(* IEC 61131-3 sources: PortalRobot/Portal_robot/Device/application/FB (part 2) *)

(* ---- FB_AXIS_GROUP.st ---- *)
FUNCTION_BLOCK FB_AXIS_GROUP
VAR_INPUT
	FaultRequest : ST_AXIS_GROUP_FAULT_REQUEST; // Единый контракт диагностической инъекции
	xResetPermit : BOOL; // Общий сброс разрешён ручным режимом и остановленной ячейкой
	xAxesPowered : BOOL; // Питанием физических осей владеют FB_AXIS; группа только наблюдает готовность
	lrVelocityOverride : LREAL; // Live override скорости групповых движений, 0.001..1.0
END_VAR
VAR_OUTPUT
	FaultStatus : ST_FAULT_INJECTION_STATUS; // Состояние инжектора для HMI
END_VAR
VAR
	// Внутренние исполняемые булевые переменные
	xEnable      : BOOL; // Импульс включения группы
	xDisable     : BOOL; // Импульс отключения группы
	xReset       : BOOL; // Импульс сброса ошибок
	xResetMC     : BOOL; // Выполняется сброс SoftMotion
	xMoveDirect  : BOOL; // Выполняется прямое перемещение
	xMoveLinear  : BOOL; // Выполняется линейное перемещение
	xStopCmd     : BOOL; // Выполняется остановка
	xHaltCmd     : BOOL; // Выполняется плавная остановка
	lrAppliedVelocityOverride : LREAL; // Коэффициент после защитного ограничения PLC
	xVelocityOverrideEnable : BOOL; // Запись live override разрешена только в рабочих состояниях без MC_GroupStop
	xFaultAllowed : BOOL; // Безопасные условия тестового запуска

	iPrevStep : E_AXIS_GROUP_STATE; // Предыдущий шаг автомата

	// Для таймера шага
	tonStepTimeout   : TON; // Таймер превышения времени шага
	xStepTimeout     : BOOL; // Время шага превышено
	xStepChanged     : BOOL; // Шаг изменился в текущем цикле
	xStepTimerEnable : BOOL; // Разрешение таймера шага
	xStepInitialized : BOOL; // Предыдущий шаг инициализирован

	// Для удержания предупреждений
    tpWarningHold : TP; // Удержание предупреждения для отображения
    xWarningPulse : BOOL; // Импульс нового предупреждения

	// ФБ группы осей
	fbReadStatus   : MC_GroupReadStatus; // Чтение состояния группы
	fbReadError    : MC_GroupReadError; // Чтение активной ошибки группы
	fbReadPosition : MC_GroupReadActualPosition; // Чтение текущей позиции группы
	fbGroupEnable  : MC_GroupEnable; // Включение группы
	fbGroupDisable : MC_GroupDisable; // Отключение группы
	fbGroupReset   : MC_GroupReset; // Сброс ошибок группы
	fbGroupSetOverride : MC_GroupSetOverride; // Live override активного и следующего движения группы

	fbMoveDirect : MC_MoveDirectAbsolute; // Прямое абсолютное перемещение
	fbMoveLinear : MC_MoveLinearAbsolute; // Линейное абсолютное перемещение
	fbFaultInjector : FB_AXIS_GROUP_FAULT_INJECTOR; // Изолированная инъекция библиотечной ошибки

	fbGroupHalt : MC_GroupHalt; // Плавная остановка группы
	fbGroupStop : MC_GroupStop; // Остановка группы

	stPosition : SMC_POS_REF; // Текущая позиция группы

	// Триггеры на команды
    rtEnable        : R_TRIG; // Фронт команды включения
    rtDisable       : R_TRIG; // Фронт команды отключения
	rtEnablePower   : R_TRIG; // Фронт запроса питания
    rtResetAllError : R_TRIG; // Фронт команды сброса
    rtMoveDirect    : R_TRIG; // Фронт прямого перемещения
    rtMoveLinear    : R_TRIG; // Фронт линейного перемещения
	rtStopCmd       : R_TRIG; // Фронт команды остановки
	rtHaltCmd       : R_TRIG; // Фронт плавной остановки

END_VAR
VAR_IN_OUT
	AxisGroup : AXIS_GROUP_REF_SM3; // Ссылка на группу осей SoftMotion
	GroupData : ST_AXIS_GROUP; // Команды, статусы и диагностика группы
END_VAR

VAR CONSTANT
	// ==================================================
    // Логические ошибки группы
    // ==================================================
	LOG_STEP_TIMEOUT             : DWORD := 1; // Превышено время шага
	LOG_INVALID_STATE            : DWORD := 2; // Неизвестный шаг автомата
	LOG_POWER_PERMIT_READY       : DWORD := 4; // Нет разрешения питания в готовности
	LOG_POWER_PERMIT_LOST_DIRECT : DWORD := 8; // Разрешение питания снято при движении
	// ==================================================
    // Ошибки блоков движения группы
    // ==================================================
	MOTION_ERR_ENABLE        : DWORD := 1; // Ошибка включения группы
	MOTION_ERR_DISABLE       : DWORD := 4; // Ошибка отключения группы
	MOTION_ERR_RESET         : DWORD := 8; // Ошибка сброса группы
	MOTION_ERR_MOVE_DIRECT   : DWORD := 16; // Ошибка прямого перемещения
	MOTION_ERR_MOVE_LINEAR   : DWORD := 32; // Ошибка линейного перемещения
	MOTION_ERR_HALT          : DWORD := 64; // Ошибка плавной остановки
	MOTION_ERR_STOP          : DWORD := 128; // Ошибка остановки
	MOTION_ERR_READ_POSITION : DWORD := 256; // Ошибка чтения позиции
	MOTION_ERR_READ_STATUS   : DWORD := 512; // Ошибка чтения статуса
	MOTION_ERR_READ_GROUP_ERROR : DWORD := 1024; // Ошибка чтения кода ошибки группы
	MOTION_ERR_GROUP_ERROR_STOP : DWORD := 2048; // Группа SoftMotion находится в ErrorStop
	MOTION_ERR_SIMULATED        : DWORD := 4096; // Тестовая ошибка MC_MoveDirectAbsolute
	MOTION_ERR_OVERRIDE         : DWORD := 8192; // Ошибка MC_GroupSetOverride; бит 1 сохранён за legacy POWER_ERROR

	WRN_NO_POWER_PERMIT       : UINT := 1; // Нет разрешения питания
	WRN_MOVE_COMMAND_CONFLICT : UINT := 2; // Одновременно заданы два типа движения
	WRN_GLOBAL_ERROR_ACTIVE   : UINT := 3; // Сброс отклонён из-за глобальной ошибки
	WRN_MOTION_ERROR_ACTIVE   : UINT := 4; // Сброс отклонён из-за активной Motion-ошибки
	WRN_RESET_VERIFY_TIMEOUT  : UINT := 5; // Не получено подтверждение сброса за допустимое время
	WRN_GROUP_ERROR_AFTER_RESET : UINT := 6; // Группа осталась в ErrorStop после сброса
	WRN_GROUP_RESET_ERROR     : UINT := 7; // MC_GroupReset завершился ошибкой
	WRN_GROUP_RESET_TIMEOUT   : UINT := 8; // Превышено время выполнения MC_GroupReset
	WRN_SIM_ERROR_NOT_ALLOWED : UINT := 9; // Тестовая ошибка запрещена текущим состоянием группы
END_VAR

// --- BEGIN IMPLEMENTATION ---

// Коэффициент симуляции не изменяет динамику группы осей робота.
lrAppliedVelocityOverride := MAX(0.001, MIN(1.0, lrVelocityOverride));

// =============================================================================
// 1. Добить предупреждения и ошибки
// 2. Сделать логирование ошибок и шагов
// 3. Сделать необходимые сигналы статусов
// =============================================================================

// =============================================================================
// 1. Одноцикловые сигналы
// =============================================================================
xWarningPulse := FALSE;

GroupData.Diag.xStepChanged := FALSE;
GroupData.Error.dwLogicalErrorNew := DWORD#0;
GroupData.Error.dwMotionErrorNew := DWORD#0;

// =============================================================================
// 2. Фронты команд
// =============================================================================
rtDisable(CLK := GroupData.Command.xDisable);
rtEnablePower(CLK := GroupData.Command.xPowerEnable);
rtResetAllError(CLK := GroupData.Command.xReset);
rtMoveDirect(CLK := GroupData.Command.xMoveDirect);
rtMoveLinear(CLK := GroupData.Command.xMoveLinear);
rtHaltCmd(CLK := GroupData.Command.xHaltCmd);
rtStopCmd(CLK := GroupData.Command.xStopCmd);

// =============================================================================
// 3. Чтение состояния группы и координат
// =============================================================================
fbReadStatus(
    Enable    := TRUE,
    AxisGroup := AxisGroup
);

fbReadError(
    Enable    := TRUE,
    AxisGroup := AxisGroup
);

fbReadPosition(
    AxisGroup   := AxisGroup,
    Enable      := TRUE,
    CoordSystem := SMC_COORD_SYSTEM.MCS
);

IF fbReadPosition.Valid THEN
	stPosition := fbReadPosition.Position;
    GroupData.Status.ActualX := fbReadPosition.Position.c.X;
    GroupData.Status.ActualY := fbReadPosition.Position.c.Y;
    GroupData.Status.ActualZ := fbReadPosition.Position.c.Z;
END_IF;
GroupData.Status.xPositionValid := fbReadPosition.Valid AND NOT fbReadPosition.Error;

// =============================================================================
// 4. Текущий статус ошибок
// =============================================================================
GroupData.Status.xGroupError :=
    fbReadStatus.Error
    OR fbReadStatus.GroupErrorStop
    OR (GroupData.Error.dwMotionErrorLatched <> DWORD#0);

GroupData.Status.xLogicalError :=
    GroupData.Error.dwLogicalErrorLatched <> DWORD#0;

GroupData.Status.xLocalError :=
    GroupData.Status.xGroupError
    OR GroupData.Status.xLogicalError;

// Тестовый Motion-FB запускается только в неподвижной готовой группе.
xFaultAllowed := fbReadStatus.Valid
	AND fbReadStatus.GroupStandby
	AND (GroupData.Diag.iStep = E_AXIS_GROUP_STATE.READY)
	AND NOT GroupData.Status.xLocalError
	AND NOT GroupData.Command.xGlobalError
	AND NOT GroupData.Command.xMoveDirect
	AND NOT GroupData.Command.xMoveLinear;

fbFaultInjector(
	Request := FaultRequest,
	xOwnerAllowed := xFaultAllowed,
	xReset := GroupData.Command.xReset,
	Position := stPosition,
	AxisGroup := AxisGroup
);
FaultStatus := fbFaultInjector.Status;

IF fbFaultInjector.Status.xRejected THEN
	GroupData.Diag.sWarningText := 'Simulated SM3 error is not allowed';
	GroupData.Diag.stWarning.uiCode := WRN_SIM_ERROR_NOT_ALLOWED;
	GroupData.Diag.stWarning.udiSequence := GroupData.Diag.stWarning.udiSequence + UDINT#1;
	IF GroupData.Diag.stWarning.udiSequence = UDINT#0 THEN
		GroupData.Diag.stWarning.udiSequence := UDINT#1;
	END_IF;
	xWarningPulse := TRUE;
END_IF;

// =============================================================================
// 5. Команды Motion FB по умолчанию
// =============================================================================
xEnable := FALSE;
xDisable := FALSE;
xResetMC := FALSE;
xMoveDirect := FALSE;
xMoveLinear := FALSE;
xStopCmd := FALSE;
xHaltCmd := FALSE;

// =============================================================================
// 6. Машина состояний
// =============================================================================
CASE GroupData.Diag.iStep OF

    // -------------------------------------------------------------------------
    E_AXIS_GROUP_STATE.DISABLED:
    // -------------------------------------------------------------------------
        GroupData.Diag.sStepName := 'DISABLED';
        GroupData.Diag.tStepPreset := T#0S;
        GroupData.Diag.iPowerMode := E_AXIS_GROUP_POWER_MODE.OFF;

        IF GroupData.Command.xGlobalError
           OR GroupData.Status.xLocalError THEN

            GroupData.Diag.iStep := E_AXIS_GROUP_STATE.ERROR;

        ELSIF rtEnablePower.Q AND NOT GroupData.Command.xPowerPermit THEN
            GroupData.Diag.sWarningText := 'Power permit is not active';
            GroupData.Diag.stWarning.uiCode := WRN_NO_POWER_PERMIT;
            GroupData.Diag.stWarning.udiSequence := GroupData.Diag.stWarning.udiSequence + UDINT#1;
            IF GroupData.Diag.stWarning.udiSequence = UDINT#0 THEN
                GroupData.Diag.stWarning.udiSequence := UDINT#1;
            END_IF;
            xWarningPulse := TRUE;

		ELSIF fbReadStatus.Valid AND fbReadStatus.GroupStandby THEN
			// MC_GroupReset всегда возвращает группу в GroupStandby. Если питание
			// запрошено, используем это состояние без повторного MC_GroupEnable;
			// иначе сначала синхронизируем группу с программным шагом DISABLED.
			IF rtEnablePower.Q THEN
				GroupData.Diag.iStep := E_AXIS_GROUP_STATE.ENABLING_POWER;
			ELSE
				GroupData.Diag.iStep := E_AXIS_GROUP_STATE.DISABLING_GROUP;
			END_IF;

        ELSIF rtEnablePower.Q THEN
            GroupData.Diag.iStep := E_AXIS_GROUP_STATE.ENABLING_POWER;
        END_IF;

    // -------------------------------------------------------------------------
    E_AXIS_GROUP_STATE.ENABLING_POWER:
    // -------------------------------------------------------------------------
        GroupData.Diag.sStepName := 'ENABLING_POWER';
        GroupData.Diag.tStepPreset := GroupData.Timeouts.tPowerTimeout;
        GroupData.Diag.iPowerMode := E_AXIS_GROUP_POWER_MODE.ON;

        IF fbReadStatus.GroupErrorStop THEN

            GroupData.Diag.iStep := E_AXIS_GROUP_STATE.ERROR;

        ELSIF NOT GroupData.Command.xPowerPermit
           OR GroupData.Command.xGlobalError THEN

            GroupData.Diag.iStep := E_AXIS_GROUP_STATE.DISABLING_POWER;

        ELSIF xStepTimeout THEN
            GroupData.Error.dwLogicalErrorNew :=
                GroupData.Error.dwLogicalErrorNew
                OR LOG_STEP_TIMEOUT;

            GroupData.Diag.iStep := E_AXIS_GROUP_STATE.DISABLING_POWER;

		ELSIF xAxesPowered AND fbReadStatus.Valid THEN
			IF fbReadStatus.GroupStandby THEN
				GroupData.Diag.iStep := E_AXIS_GROUP_STATE.READY;
			ELSIF fbReadStatus.GroupDisabled THEN
				GroupData.Diag.iStep := E_AXIS_GROUP_STATE.ENABLING_GROUP;
			END_IF;
		END_IF;

    // -------------------------------------------------------------------------
    E_AXIS_GROUP_STATE.ENABLING_GROUP:
    // -------------------------------------------------------------------------
        GroupData.Diag.sStepName := 'ENABLING_GROUP';
        GroupData.Diag.tStepPreset := GroupData.Timeouts.tGroupTimeout;
        GroupData.Diag.iPowerMode := E_AXIS_GROUP_POWER_MODE.ON;

		// MC_GroupEnable допустим только из GroupDisabled. Execute формируется
		// исключительно на этом шаге: после перехода в GroupStandby он снимается,
		// чтобы новый фронт не вызвал MC_GroupEnable повторно после MC_GroupReset.
		xEnable := fbReadStatus.Valid AND fbReadStatus.GroupDisabled;

		IF fbReadStatus.GroupErrorStop THEN

            GroupData.Diag.iStep := E_AXIS_GROUP_STATE.ERROR;

		ELSIF fbReadStatus.Valid AND fbReadStatus.GroupStandby THEN

			GroupData.Diag.iStep := E_AXIS_GROUP_STATE.READY;

		ELSIF xEnable AND fbGroupEnable.Error THEN

			GroupData.Diag.iStep := E_AXIS_GROUP_STATE.ERROR;

        ELSIF NOT GroupData.Command.xPowerPermit
           OR GroupData.Command.xGlobalError THEN

            GroupData.Diag.iStep := E_AXIS_GROUP_STATE.DISABLING_GROUP;

        ELSIF xStepTimeout THEN
            GroupData.Error.dwLogicalErrorNew :=
                GroupData.Error.dwLogicalErrorNew
                OR LOG_STEP_TIMEOUT;

            GroupData.Diag.iStep := E_AXIS_GROUP_STATE.DISABLING_GROUP;

		END_IF;

    // -------------------------------------------------------------------------
    E_AXIS_GROUP_STATE.READY:
    // -------------------------------------------------------------------------
        GroupData.Diag.sStepName := 'READY';
        GroupData.Diag.tStepPreset := T#0S;
        GroupData.Diag.iPowerMode := E_AXIS_GROUP_POWER_MODE.ON;

		IF fbReadStatus.GroupErrorStop THEN
            GroupData.Diag.iStep := E_AXIS_GROUP_STATE.ERROR;

        ELSIF NOT GroupData.Command.xPowerPermit
           OR GroupData.Command.xGlobalError
           OR GroupData.Status.xLocalError
           OR rtDisable.Q THEN

            GroupData.Diag.iStep := E_AXIS_GROUP_STATE.DISABLING_GROUP;

        ELSIF rtMoveDirect.Q AND rtMoveLinear.Q THEN
            GroupData.Diag.sWarningText :=
                'MoveDirect and MoveLinear requested together';

            GroupData.Diag.stWarning.uiCode := WRN_MOVE_COMMAND_CONFLICT;
            GroupData.Diag.stWarning.udiSequence := GroupData.Diag.stWarning.udiSequence + UDINT#1;
            IF GroupData.Diag.stWarning.udiSequence = UDINT#0 THEN
                GroupData.Diag.stWarning.udiSequence := UDINT#1;
            END_IF;

            xWarningPulse := TRUE;

        ELSIF rtMoveDirect.Q THEN
            GroupData.Diag.iStep := E_AXIS_GROUP_STATE.MOVING_DIRECT;

        ELSIF rtMoveLinear.Q THEN
            GroupData.Diag.iStep := E_AXIS_GROUP_STATE.MOVING_LINEAR;
        END_IF;

    // -------------------------------------------------------------------------
    E_AXIS_GROUP_STATE.MOVING_DIRECT:
    // -------------------------------------------------------------------------
        GroupData.Diag.sStepName := 'MOVING_DIRECT';
        GroupData.Diag.tStepPreset := GroupData.Timeouts.tMoveTimeout;
        GroupData.Diag.iPowerMode := E_AXIS_GROUP_POWER_MODE.ON;

		xMoveDirect := TRUE;

        IF fbReadStatus.GroupErrorStop THEN
            GroupData.Diag.iStep := E_AXIS_GROUP_STATE.ERROR;

        ELSIF fbMoveDirect.Error THEN
            IF fbReadStatus.GroupMoving THEN
                GroupData.Diag.iStep := E_AXIS_GROUP_STATE.EMG_STOP;
            ELSE
                GroupData.Diag.iStep := E_AXIS_GROUP_STATE.ERROR;
            END_IF;

        ELSIF xStepTimeout THEN
            GroupData.Error.dwLogicalErrorNew :=
                GroupData.Error.dwLogicalErrorNew
                OR LOG_STEP_TIMEOUT;

            GroupData.Diag.iStep := E_AXIS_GROUP_STATE.EMG_STOP;

        ELSIF NOT GroupData.Command.xPowerPermit
           OR GroupData.Command.xGlobalError
           OR GroupData.Status.xLocalError
           OR rtStopCmd.Q THEN

            GroupData.Diag.iStep := E_AXIS_GROUP_STATE.EMG_STOP;

        ELSIF rtHaltCmd.Q THEN
            GroupData.Diag.iStep := E_AXIS_GROUP_STATE.HALT_STOP;

        ELSIF fbMoveDirect.Done
           AND fbReadStatus.GroupStandby THEN

            GroupData.Diag.iStep := E_AXIS_GROUP_STATE.READY;
        END_IF;

    // -------------------------------------------------------------------------
    E_AXIS_GROUP_STATE.HALT_STOP:
    // -------------------------------------------------------------------------
        GroupData.Diag.sStepName := 'HALT_STOP';
        GroupData.Diag.tStepPreset := GroupData.Timeouts.tHaltTimeout;
        GroupData.Diag.iPowerMode := E_AXIS_GROUP_POWER_MODE.ON;

		xHaltCmd := TRUE;

        IF fbReadStatus.GroupErrorStop THEN
            GroupData.Diag.iStep := E_AXIS_GROUP_STATE.ERROR;

        ELSIF fbGroupHalt.Error
           OR xStepTimeout
           OR NOT GroupData.Command.xPowerPermit
           OR GroupData.Command.xGlobalError
           OR GroupData.Status.xLocalError
           OR rtStopCmd.Q THEN

            IF xStepTimeout THEN
                GroupData.Error.dwLogicalErrorNew :=
                    GroupData.Error.dwLogicalErrorNew
                    OR LOG_STEP_TIMEOUT;
            END_IF;

            GroupData.Diag.iStep := E_AXIS_GROUP_STATE.EMG_STOP;

        ELSIF fbGroupHalt.Done
           AND fbReadStatus.GroupStandby THEN

            GroupData.Diag.iStep := E_AXIS_GROUP_STATE.READY;
        END_IF;

    // -------------------------------------------------------------------------
    E_AXIS_GROUP_STATE.EMG_STOP:
    // -------------------------------------------------------------------------
        GroupData.Diag.sStepName := 'STOPPING';
        GroupData.Diag.tStepPreset := GroupData.Timeouts.tStopTimeout;
        GroupData.Diag.iPowerMode := E_AXIS_GROUP_POWER_MODE.ON;

		xStopCmd := TRUE;

        IF fbReadStatus.GroupErrorStop
           OR fbGroupStop.Error THEN

            GroupData.Diag.iStep := E_AXIS_GROUP_STATE.ERROR;

        ELSIF xStepTimeout THEN
            GroupData.Error.dwLogicalErrorNew :=
                GroupData.Error.dwLogicalErrorNew
                OR LOG_STEP_TIMEOUT;

            GroupData.Diag.iStep := E_AXIS_GROUP_STATE.ERROR;

        ELSIF fbGroupStop.Done THEN
            GroupData.Diag.iStep := E_AXIS_GROUP_STATE.WAIT_STOP;
        END_IF;

    // -------------------------------------------------------------------------
    E_AXIS_GROUP_STATE.WAIT_STOP:
    // -------------------------------------------------------------------------
        GroupData.Diag.sStepName := 'WAIT_STOP';
        GroupData.Diag.tStepPreset := GroupData.Timeouts.tStopTimeout;
        GroupData.Diag.iPowerMode := E_AXIS_GROUP_POWER_MODE.ON;

		IF fbReadStatus.GroupErrorStop THEN
            GroupData.Diag.iStep := E_AXIS_GROUP_STATE.ERROR;

        ELSIF xStepTimeout THEN
            GroupData.Error.dwLogicalErrorNew :=
                GroupData.Error.dwLogicalErrorNew
                OR LOG_STEP_TIMEOUT;

            GroupData.Diag.iStep := E_AXIS_GROUP_STATE.ERROR;

		ELSIF fbReadStatus.GroupStandby THEN
			// Операторский Stop завершает только движение и сохраняет GroupStandby.
			// Отключение группы выполняется лишь по отдельному запросу питания/ошибке.
			IF GroupData.Command.xPowerPermit
			AND NOT GroupData.Command.xDisable
			AND NOT GroupData.Command.xGlobalError
			AND NOT GroupData.Status.xLocalError THEN
				GroupData.Diag.iStep := E_AXIS_GROUP_STATE.READY;
			ELSE
				GroupData.Diag.iStep := E_AXIS_GROUP_STATE.DISABLING_GROUP;
			END_IF;
		END_IF;

    // -------------------------------------------------------------------------
    E_AXIS_GROUP_STATE.DISABLING_GROUP:
    // -------------------------------------------------------------------------
        GroupData.Diag.sStepName := 'DISABLING_GROUP';
        GroupData.Diag.tStepPreset := GroupData.Timeouts.tGroupTimeout;
        GroupData.Diag.iPowerMode := E_AXIS_GROUP_POWER_MODE.ON;

		// MC_GroupDisable допустим только из GroupStandby.
		xDisable := fbReadStatus.Valid AND fbReadStatus.GroupStandby;

		IF fbReadStatus.GroupErrorStop THEN

            GroupData.Diag.iStep := E_AXIS_GROUP_STATE.ERROR;

		ELSIF fbReadStatus.Valid AND fbReadStatus.GroupDisabled THEN

			GroupData.Diag.iStep := E_AXIS_GROUP_STATE.DISABLING_POWER;

		ELSIF xDisable AND fbGroupDisable.Error THEN

			GroupData.Diag.iStep := E_AXIS_GROUP_STATE.ERROR;

        ELSIF xStepTimeout THEN
            GroupData.Error.dwLogicalErrorNew :=
                GroupData.Error.dwLogicalErrorNew
                OR LOG_STEP_TIMEOUT;

            GroupData.Diag.iStep := E_AXIS_GROUP_STATE.ERROR;

		ELSIF xDisable AND fbGroupDisable.Done
           AND fbReadStatus.GroupDisabled THEN

            GroupData.Diag.iStep := E_AXIS_GROUP_STATE.DISABLING_POWER;
        END_IF;

    // -------------------------------------------------------------------------
    E_AXIS_GROUP_STATE.DISABLING_POWER:
    // -------------------------------------------------------------------------
        GroupData.Diag.sStepName := 'DISABLING_POWER';
        GroupData.Diag.tStepPreset := GroupData.Timeouts.tPowerTimeout;
        GroupData.Diag.iPowerMode :=
            E_AXIS_GROUP_POWER_MODE.OFF_REQUEST;

        IF xStepTimeout THEN
            GroupData.Error.dwLogicalErrorNew :=
                GroupData.Error.dwLogicalErrorNew
                OR LOG_STEP_TIMEOUT;

            GroupData.Diag.iStep := E_AXIS_GROUP_STATE.ERROR;

        ELSIF NOT xAxesPowered THEN

            IF GroupData.Command.xGlobalError
               OR GroupData.Status.xLocalError
			   OR NOT GroupData.Command.xPowerPermit THEN

                GroupData.Diag.iStep := E_AXIS_GROUP_STATE.ERROR;
            ELSE
                GroupData.Diag.iStep := E_AXIS_GROUP_STATE.DISABLED;
            END_IF;
        END_IF;

    // -------------------------------------------------------------------------
    E_AXIS_GROUP_STATE.ERROR:
    // -------------------------------------------------------------------------
        GroupData.Diag.sStepName := 'ERROR';
        GroupData.Diag.tStepPreset := T#0S;

        GroupData.Diag.iPowerMode := E_AXIS_GROUP_POWER_MODE.OFF_REQUEST;

		IF rtResetAllError.Q AND xResetPermit THEN

            IF GroupData.Command.xGlobalError THEN
                GroupData.Diag.sWarningText :=
                    'Global error is still active';

                GroupData.Diag.stWarning.uiCode := WRN_GLOBAL_ERROR_ACTIVE;
                GroupData.Diag.stWarning.udiSequence := GroupData.Diag.stWarning.udiSequence + UDINT#1;
                IF GroupData.Diag.stWarning.udiSequence = UDINT#0 THEN
                    GroupData.Diag.stWarning.udiSequence := UDINT#1;
                END_IF;

                xWarningPulse := TRUE;

            ELSIF fbReadStatus.GroupErrorStop THEN
                    GroupData.Diag.iStep :=
                        E_AXIS_GROUP_STATE.RESETTING;

            ELSIF GroupData.Error.dwMotionErrorActive
                  <> DWORD#0 THEN

                GroupData.Diag.sWarningText :=
                    'Motion FB error is still active';

                GroupData.Diag.stWarning.uiCode := WRN_MOTION_ERROR_ACTIVE;
                GroupData.Diag.stWarning.udiSequence := GroupData.Diag.stWarning.udiSequence + UDINT#1;
                IF GroupData.Diag.stWarning.udiSequence = UDINT#0 THEN
                    GroupData.Diag.stWarning.udiSequence := UDINT#1;
                END_IF;

                xWarningPulse := TRUE;

            ELSE
                // Ошибка устранена — очищаем защёлки.
                GroupData.Error.dwLogicalErrorLatched := DWORD#0;
                GroupData.Error.dwMotionErrorLatched := DWORD#0;
                GroupData.Error.dwMotionErrorPrevious := DWORD#0;

				IF fbReadStatus.GroupStandby AND NOT xAxesPowered THEN
					GroupData.Diag.iStep :=
						E_AXIS_GROUP_STATE.DISABLING_GROUP;

				ELSIF fbReadStatus.GroupDisabled AND NOT xAxesPowered THEN
					GroupData.Diag.iStep :=
						E_AXIS_GROUP_STATE.DISABLED;

				ELSIF fbReadStatus.GroupDisabled THEN
					GroupData.Diag.iStep :=
						E_AXIS_GROUP_STATE.ENABLING_GROUP;

                ELSIF fbReadStatus.GroupStandby THEN
                    GroupData.Diag.iStep :=
                        E_AXIS_GROUP_STATE.READY;

                ELSE
                    GroupData.Diag.iStep :=
                        E_AXIS_GROUP_STATE.DISABLING_POWER;
                END_IF;
            END_IF;
        END_IF;

    // -------------------------------------------------------------------------
    E_AXIS_GROUP_STATE.RESETTING:
    // -------------------------------------------------------------------------
        GroupData.Diag.sStepName := 'RESETTING';
        GroupData.Diag.tStepPreset := GroupData.Timeouts.tGroupTimeout;
        GroupData.Diag.iPowerMode := E_AXIS_GROUP_POWER_MODE.ON;

		// Ошибка оси могла исчезнуть между принятием общей команды и этим циклом.
		// В таком случае MC_GroupReset не вызывается, иначе он вернёт 78
		// (no error to be resetted); остаётся только очистить внутренние защёлки.
		IF fbReadStatus.Valid AND NOT fbReadStatus.GroupErrorStop THEN
			xResetMC := FALSE;
			GroupData.Diag.iStep := E_AXIS_GROUP_STATE.RESET_VERIFY;

		ELSE
			xResetMC := TRUE;
		END_IF;

		IF GroupData.Command.xGlobalError THEN
            GroupData.Diag.sWarningText :=
                'Global error became active during group reset';

            GroupData.Diag.stWarning.uiCode := WRN_GLOBAL_ERROR_ACTIVE;
            GroupData.Diag.stWarning.udiSequence := GroupData.Diag.stWarning.udiSequence + UDINT#1;
            IF GroupData.Diag.stWarning.udiSequence = UDINT#0 THEN
                GroupData.Diag.stWarning.udiSequence := UDINT#1;
            END_IF;

            xWarningPulse := TRUE;
            GroupData.Diag.iStep := E_AXIS_GROUP_STATE.ERROR;

		ELSIF xResetMC AND fbGroupReset.Error THEN
            GroupData.Diag.sWarningText :=
                'MC_GroupReset finished with error';

            GroupData.Diag.stWarning.uiCode := WRN_GROUP_RESET_ERROR;
            GroupData.Diag.stWarning.udiSequence := GroupData.Diag.stWarning.udiSequence + UDINT#1;
            IF GroupData.Diag.stWarning.udiSequence = UDINT#0 THEN
                GroupData.Diag.stWarning.udiSequence := UDINT#1;
            END_IF;

            xWarningPulse := TRUE;
            GroupData.Diag.iStep := E_AXIS_GROUP_STATE.ERROR;

		ELSIF xResetMC AND xStepTimeout THEN
            GroupData.Diag.sWarningText :=
                'MC_GroupReset timeout';

            GroupData.Diag.stWarning.uiCode := WRN_GROUP_RESET_TIMEOUT;
            GroupData.Diag.stWarning.udiSequence := GroupData.Diag.stWarning.udiSequence + UDINT#1;
            IF GroupData.Diag.stWarning.udiSequence = UDINT#0 THEN
                GroupData.Diag.stWarning.udiSequence := UDINT#1;
            END_IF;

            xWarningPulse := TRUE;
            GroupData.Error.dwLogicalErrorNew :=
                GroupData.Error.dwLogicalErrorNew
                OR LOG_STEP_TIMEOUT;

            GroupData.Diag.iStep := E_AXIS_GROUP_STATE.ERROR;

		ELSIF xResetMC AND fbGroupReset.Done THEN
            // Статус группы был прочитан до вызова MC_GroupReset.
            // Проверяем результат сброса только со следующего цикла.
            GroupData.Diag.iStep := E_AXIS_GROUP_STATE.RESET_VERIFY;
        END_IF;

    // -------------------------------------------------------------------------
    E_AXIS_GROUP_STATE.RESET_VERIFY:
    // -------------------------------------------------------------------------
        GroupData.Diag.sStepName := 'RESET_VERIFY';
        GroupData.Diag.tStepPreset := GroupData.Timeouts.tGroupTimeout;
        GroupData.Diag.iPowerMode := E_AXIS_GROUP_POWER_MODE.ON;

        IF GroupData.Command.xGlobalError THEN
            GroupData.Diag.sWarningText :=
                'Global error became active during reset verification';

            GroupData.Diag.stWarning.uiCode := WRN_GLOBAL_ERROR_ACTIVE;
            GroupData.Diag.stWarning.udiSequence := GroupData.Diag.stWarning.udiSequence + UDINT#1;
            IF GroupData.Diag.stWarning.udiSequence = UDINT#0 THEN
                GroupData.Diag.stWarning.udiSequence := UDINT#1;
            END_IF;

            xWarningPulse := TRUE;
            GroupData.Diag.iStep := E_AXIS_GROUP_STATE.ERROR;

        ELSIF xStepTimeout THEN
            GroupData.Diag.sWarningText :=
                'Reset verification timeout';

            GroupData.Diag.stWarning.uiCode := WRN_RESET_VERIFY_TIMEOUT;
            GroupData.Diag.stWarning.udiSequence := GroupData.Diag.stWarning.udiSequence + UDINT#1;
            IF GroupData.Diag.stWarning.udiSequence = UDINT#0 THEN
                GroupData.Diag.stWarning.udiSequence := UDINT#1;
            END_IF;

            xWarningPulse := TRUE;
            GroupData.Error.dwLogicalErrorNew :=
                GroupData.Error.dwLogicalErrorNew
                OR LOG_STEP_TIMEOUT;

            GroupData.Diag.iStep := E_AXIS_GROUP_STATE.ERROR;

        ELSIF fbReadStatus.Valid
           AND fbReadStatus.GroupErrorStop
           AND fbReadError.Valid
           AND (TO_UDINT(fbReadError.GroupErrorID) <> UDINT#0) THEN

            // Причина ошибки осталась активной после завершения сброса.
            GroupData.Diag.sWarningText :=
                'Axis group error remains active after reset';

            GroupData.Diag.stWarning.uiCode := WRN_GROUP_ERROR_AFTER_RESET;
            GroupData.Diag.stWarning.udiSequence := GroupData.Diag.stWarning.udiSequence + UDINT#1;
            IF GroupData.Diag.stWarning.udiSequence = UDINT#0 THEN
                GroupData.Diag.stWarning.udiSequence := UDINT#1;
            END_IF;

            xWarningPulse := TRUE;
            GroupData.Diag.iStep := E_AXIS_GROUP_STATE.ERROR;

        ELSIF fbReadStatus.Valid
           AND NOT fbReadStatus.GroupErrorStop THEN

            GroupData.Error.dwLogicalErrorLatched := DWORD#0;
            GroupData.Error.dwMotionErrorLatched := DWORD#0;
            GroupData.Error.dwMotionErrorPrevious := DWORD#0;

			IF fbReadStatus.GroupStandby AND NOT xAxesPowered THEN
				GroupData.Diag.iStep := E_AXIS_GROUP_STATE.DISABLING_GROUP;

			ELSIF fbReadStatus.GroupDisabled AND NOT xAxesPowered THEN
				GroupData.Diag.iStep := E_AXIS_GROUP_STATE.DISABLED;

			ELSIF fbReadStatus.GroupDisabled THEN
				GroupData.Diag.iStep := E_AXIS_GROUP_STATE.ENABLING_GROUP;

            ELSIF fbReadStatus.GroupStandby THEN
                GroupData.Diag.iStep := E_AXIS_GROUP_STATE.READY;

            ELSE
                GroupData.Diag.iStep := E_AXIS_GROUP_STATE.DISABLING_POWER;
            END_IF;
        END_IF;

    // -------------------------------------------------------------------------
    ELSE
    // -------------------------------------------------------------------------
        GroupData.Error.dwLogicalErrorNew :=
            GroupData.Error.dwLogicalErrorNew
            OR LOG_INVALID_STATE;

        GroupData.Diag.iStep := E_AXIS_GROUP_STATE.ERROR;

END_CASE;

// =============================================================================
// 7. Целевая позиция
// =============================================================================
GroupData.MotionParam.stTargetPos.c.X := GroupData.MotionParam.lrX;
GroupData.MotionParam.stTargetPos.c.Y := GroupData.MotionParam.lrY;
GroupData.MotionParam.stTargetPos.c.Z := GroupData.MotionParam.lrZ;

// =============================================================================
// 8. Вызовы Motion FB
// =============================================================================
fbGroupEnable(
    AxisGroup := AxisGroup,
    Execute   := xEnable
);

fbGroupDisable(
    AxisGroup := AxisGroup,
    Execute   := xDisable
);

fbGroupReset(
    AxisGroup := AxisGroup,
    Execute   := xResetMC
);

// MC_GroupSetOverride меняет скорость уже активного движения. Вызов обязан
// находиться перед Motion FB. Во время MC_GroupStop блок запрещён документацией:
// последняя записанная величина сохраняется, а Stop выполняется со своей динамикой.
xVelocityOverrideEnable := fbReadStatus.Valid
	AND NOT fbReadStatus.GroupErrorStop
	AND NOT xStopCmd
	AND ((GroupData.Diag.iStep = E_AXIS_GROUP_STATE.READY)
		OR (GroupData.Diag.iStep = E_AXIS_GROUP_STATE.MOVING_DIRECT)
		OR (GroupData.Diag.iStep = E_AXIS_GROUP_STATE.MOVING_LINEAR));
fbGroupSetOverride(
	AxisGroup      := AxisGroup,
	Enable         := xVelocityOverrideEnable,
	VelFactor      := lrAppliedVelocityOverride,
	AccFactor      := 1.0,
	JerkFactor     := 1.0,
	TorqueFactor   := 1.0,
	PathVelFactor  := lrAppliedVelocityOverride,
	PathAccFactor  := 1.0,
	PathJerkFactor := 1.0
);

fbMoveDirect(
    AxisGroup   := AxisGroup,
    Execute     := xMoveDirect,
    Position    := GroupData.MotionParam.stTargetPos,
    CoordSystem := SMC_COORD_SYSTEM.MCS,
    BufferMode  := MC_BUFFER_MODE.Aborting,
	// Коэффициент точки задаёт профиль команды, общий процент накладывается
	// отдельно через MC_GroupSetOverride и потому здесь повторно не умножается.
	VelFactor   := MAX(0.001, MIN(1.0, GroupData.MotionParam.VelFactor)),
    AccFactor   := GroupData.MotionParam.AccFactor,
    JerkFactor  := GroupData.MotionParam.JerkFactor
);

fbMoveLinear(
    AxisGroup := AxisGroup,
    Execute   := xMoveLinear
);

fbGroupHalt(
	AxisGroup    := AxisGroup,
	Execute      := xHaltCmd,
	Deceleration := GroupData.MotionParam.HaltDeceleration,
	Jerk         := GroupData.MotionParam.HaltJerk
);

fbGroupStop(
	AxisGroup    := AxisGroup,
	Execute      := xStopCmd,
	Deceleration := GroupData.MotionParam.HaltDeceleration * 2,
	Jerk         := GroupData.MotionParam.HaltJerk * 2
);

// =============================================================================
// 9. Маска Motion-ошибок
// =============================================================================
GroupData.Error.dwMotionErrorActive := DWORD#0;

IF fbGroupEnable.Error THEN
    GroupData.Error.dwMotionErrorActive :=
        GroupData.Error.dwMotionErrorActive
        OR MOTION_ERR_ENABLE;
END_IF;

IF fbGroupDisable.Error THEN
    GroupData.Error.dwMotionErrorActive :=
        GroupData.Error.dwMotionErrorActive
        OR MOTION_ERR_DISABLE;
END_IF;

IF fbGroupReset.Error THEN
    GroupData.Error.dwMotionErrorActive :=
        GroupData.Error.dwMotionErrorActive
        OR MOTION_ERR_RESET;
END_IF;

IF fbMoveDirect.Error THEN
    GroupData.Error.dwMotionErrorActive :=
        GroupData.Error.dwMotionErrorActive
        OR MOTION_ERR_MOVE_DIRECT;
END_IF;

IF fbMoveLinear.Error THEN
    GroupData.Error.dwMotionErrorActive :=
        GroupData.Error.dwMotionErrorActive
        OR MOTION_ERR_MOVE_LINEAR;
END_IF;

IF fbGroupHalt.Error THEN
    GroupData.Error.dwMotionErrorActive :=
        GroupData.Error.dwMotionErrorActive
        OR MOTION_ERR_HALT;
END_IF;

IF fbGroupStop.Error THEN
    GroupData.Error.dwMotionErrorActive :=
        GroupData.Error.dwMotionErrorActive
        OR MOTION_ERR_STOP;
END_IF;

IF fbReadPosition.Error THEN
    GroupData.Error.dwMotionErrorActive :=
        GroupData.Error.dwMotionErrorActive
        OR MOTION_ERR_READ_POSITION;
END_IF;

IF fbReadStatus.Error THEN
    GroupData.Error.dwMotionErrorActive :=
        GroupData.Error.dwMotionErrorActive
        OR MOTION_ERR_READ_STATUS;
END_IF;

IF fbReadError.Error THEN
    GroupData.Error.dwMotionErrorActive :=
        GroupData.Error.dwMotionErrorActive
        OR MOTION_ERR_READ_GROUP_ERROR;
END_IF;

IF fbReadStatus.GroupErrorStop THEN
    GroupData.Error.dwMotionErrorActive :=
        GroupData.Error.dwMotionErrorActive
        OR MOTION_ERR_GROUP_ERROR_STOP;
END_IF;

IF fbFaultInjector.xError THEN
	GroupData.Error.dwMotionErrorActive :=
		GroupData.Error.dwMotionErrorActive
		OR MOTION_ERR_SIMULATED;
END_IF;

IF fbGroupSetOverride.Error THEN
	GroupData.Error.dwMotionErrorActive :=
		GroupData.Error.dwMotionErrorActive
		OR MOTION_ERR_OVERRIDE;
END_IF;

// Только ошибки, которых не было в предыдущем цикле.
GroupData.Error.dwMotionErrorNew :=
    GroupData.Error.dwMotionErrorActive
    AND NOT GroupData.Error.dwMotionErrorPrevious;

// Защёлкиваем новые логические и Motion-ошибки.
GroupData.Error.dwLogicalErrorLatched :=
    GroupData.Error.dwLogicalErrorLatched
    OR GroupData.Error.dwLogicalErrorNew;

GroupData.Error.dwMotionErrorLatched :=
    GroupData.Error.dwMotionErrorLatched
    OR GroupData.Error.dwMotionErrorNew;

// Сохраняем Motion-маску для следующего цикла.
GroupData.Error.dwMotionErrorPrevious :=
    GroupData.Error.dwMotionErrorActive;

GroupData.Error.dwAlarmActive :=
    GroupData.Error.dwMotionErrorLatched
    OR SHL(GroupData.Error.dwLogicalErrorLatched, 16);

// =============================================================================
// 11. Изменение шага и таймер
// =============================================================================
IF NOT xStepInitialized THEN
    iPrevStep := GroupData.Diag.iStep;
    xStepInitialized := TRUE;
END_IF;

xStepChanged :=
    GroupData.Diag.iStep <> iPrevStep;

GroupData.Diag.xStepChanged := xStepChanged;

IF xStepChanged THEN
    GroupData.Diag.iOldStep := iPrevStep;
    GroupData.Diag.iNewStep := GroupData.Diag.iStep;
    iPrevStep := GroupData.Diag.iStep;
END_IF;

// При переходе в новый шаг таймер один цикл выключен.
// Со следующего цикла начинается отсчёт нового шага.
tonStepTimeout(
    IN :=
        NOT xStepChanged
        AND (GroupData.Diag.tStepPreset > T#0S)
        AND (GroupData.Diag.iStep <> E_AXIS_GROUP_STATE.ERROR),

    PT := GroupData.Diag.tStepPreset
);

xStepTimeout := tonStepTimeout.Q;
GroupData.Diag.xStepTimeout := xStepTimeout;

// =============================================================================
// 12. Финальные статусы
// =============================================================================
GroupData.Status.xGroupError :=
    fbReadStatus.Error
    OR fbReadStatus.GroupErrorStop
    OR (GroupData.Error.dwMotionErrorLatched <> DWORD#0);

GroupData.Status.xLogicalError :=
    GroupData.Error.dwLogicalErrorLatched <> DWORD#0;

GroupData.Status.xLocalError :=
    GroupData.Status.xGroupError
    OR GroupData.Status.xLogicalError;

GroupData.Status.xSimErrorAllowed := FaultStatus.xAllowed;

GroupData.Status.xMoveDirectDone := fbMoveDirect.Done;

// Код ошибки самой группы не совпадает с ErrorID диагностических Motion FB.
IF fbReadError.Valid
   AND (TO_UDINT(fbReadError.GroupErrorID) <> UDINT#0) THEN
    GroupData.Diag.udiActualErrorID := TO_UDINT(fbReadError.GroupErrorID);
    GroupData.Diag.sErrorText := 'Axis group error';
ELSIF (GroupData.Error.dwMotionErrorLatched AND MOTION_ERR_SIMULATED) <> DWORD#0 THEN
	GroupData.Diag.udiActualErrorID := fbFaultInjector.udiErrorID;
	GroupData.Diag.sErrorText := 'Simulated MC_MoveDirectAbsolute error';
ELSIF fbGroupSetOverride.Error THEN
	GroupData.Diag.udiActualErrorID := TO_UDINT(fbGroupSetOverride.ErrorID);
	GroupData.Diag.sErrorText := 'MC_GroupSetOverride error';
ELSIF fbGroupEnable.Error THEN
	GroupData.Diag.udiActualErrorID := TO_UDINT(fbGroupEnable.ErrorID);
	GroupData.Diag.sErrorText := 'MC_GroupEnable error';
ELSIF fbGroupDisable.Error THEN
	GroupData.Diag.udiActualErrorID := TO_UDINT(fbGroupDisable.ErrorID);
	GroupData.Diag.sErrorText := 'MC_GroupDisable error';
ELSIF fbGroupReset.Error THEN
    GroupData.Diag.udiActualErrorID := TO_UDINT(fbGroupReset.ErrorID);
    GroupData.Diag.sErrorText := 'MC_GroupReset error';
ELSIF fbMoveDirect.Error THEN
	GroupData.Diag.udiActualErrorID := TO_UDINT(fbMoveDirect.ErrorID);
	GroupData.Diag.sErrorText := 'MC_MoveDirectAbsolute error';
ELSIF fbMoveLinear.Error THEN
	GroupData.Diag.udiActualErrorID := TO_UDINT(fbMoveLinear.ErrorID);
	GroupData.Diag.sErrorText := 'MC_MoveLinearAbsolute error';
ELSIF fbGroupHalt.Error THEN
	GroupData.Diag.udiActualErrorID := TO_UDINT(fbGroupHalt.ErrorID);
	GroupData.Diag.sErrorText := 'MC_GroupHalt error';
ELSIF fbGroupStop.Error THEN
	GroupData.Diag.udiActualErrorID := TO_UDINT(fbGroupStop.ErrorID);
	GroupData.Diag.sErrorText := 'MC_GroupStop error';
ELSE
    GroupData.Diag.udiActualErrorID := UDINT#0;
    GroupData.Diag.sErrorText := '';
END_IF;

IF GroupData.Diag.udiActualErrorID <> UDINT#0 THEN
    GroupData.Diag.udiLastErrorID := GroupData.Diag.udiActualErrorID;
END_IF;

// Сохраняем последнюю ненулевую ошибку и формируем удобное представление для HMI.
IF (GroupData.Error.dwMotionErrorLatched <> DWORD#0)
OR (GroupData.Error.dwLogicalErrorLatched <> DWORD#0) THEN
	GroupData.Error.dwMotionErrorLast := GroupData.Error.dwMotionErrorLatched;
	GroupData.Error.dwLogicalErrorLast := GroupData.Error.dwLogicalErrorLatched;
END_IF;

GroupData.Error.stErrorActive := UpdateErrorView(
	dwMotionError := GroupData.Error.dwMotionErrorLatched OR GroupData.Error.dwMotionErrorActive,
	dwLogicalError := GroupData.Error.dwLogicalErrorLatched
);
GroupData.Error.stErrorLast := UpdateErrorView(
	dwMotionError := GroupData.Error.dwMotionErrorLast,
	dwLogicalError := GroupData.Error.dwLogicalErrorLast
);

// Для общей кнопки публикуется готовность владельца группы, а не только
// состояние диагностического инжектора.
FaultStatus.xResetAllowed := (GroupData.Diag.iStep = E_AXIS_GROUP_STATE.ERROR)
	AND xResetPermit
	AND NOT GroupData.Command.xGlobalError
	AND (GroupData.Status.xLocalError
		OR GroupData.Status.xLogicalError
		OR GroupData.Status.xGroupError);

(* ---- FB_CELL_SAFETY.st ---- *)
FUNCTION_BLOCK FB_CELL_SAFETY
VAR_INPUT
	axDoorLockClosedInput : ARRAY [1..4] OF BOOL;
	axDoorUnlockButtonInput : ARRAY [1..4] OF BOOL;
	axMagazineMechanismBusy : ARRAY [1..2] OF BOOL; // Только новый механизм, включая фактическое движение оси
	axEmergencyStopButtonStationInput : ARRAY [1..4] OF BOOL;
	axEmergencyStopCabinetInput : ARRAY [1..2] OF BOOL;
	xEmergencyStopMpgInput : BOOL;
	xPhaseRelayOkInput    : BOOL;
	xPressureRelayOkInput : BOOL;
	xSafetyRelayOkInput   : BOOL;
	xCellStartButtonInput : BOOL;
	xCellStopButtonInput  : BOOL;
	xCellResetButtonInput : BOOL;
	xMpgAxisXInput : BOOL;
	xMpgAxisYInput : BOOL;
	xMpgAxisZInput : BOOL;
	xMpgMultiplier1Input : BOOL;
	xMpgMultiplier10Input : BOOL;
	xMpgMultiplier100Input : BOOL;
	xSafetyRelayReset : BOOL; // Импульс отдельного сброса реле безопасности
	astMagazineStatus : ARRAY [1..2] OF ST_MAGAZINE_STATUS;
	FaultRequest : ST_CELL_SAFETY_FAULT_REQUEST;
END_VAR
VAR_OUTPUT
	Status : ST_CELL_SAFETY_STATUS;
	Error  : ST_CELL_SAFETY_ERRORS;
	Diag   : ST_CELL_SAFETY_DIAG;
	FaultStatus : ST_FAULT_INJECTION_STATUS;
	astButtonStationIoStatus : ARRAY [1..4] OF ST_BUTTON_STATION_IO_STATUS;
	stFrontControlCabinetIoStatus : ST_CONTROL_CABINET_IO_STATUS;
	stRearControlCabinetIoStatus : ST_CONTROL_CABINET_IO_STATUS;
	stMpgIoStatus : ST_MPG_IO_STATUS;
	astEnclosureDoorStatus : ARRAY [1..4] OF ST_ENCLOSURE_DOOR_STATUS;
	axDoorUnlockOutput : ARRAY [1..4] OF BOOL;
	axDoorButtonLampOutput : ARRAY [1..4] OF BOOL;
	xSafetyRelayResetOutput : BOOL;
	xCellEnablePulse : BOOL;
	xCellDisablePulse : BOOL;
	xCellResetPulse : BOOL;
END_VAR
VAR
	fbFaultInjector : FB_CELL_SAFETY_FAULT_INJECTOR;
	axEmergencyStopStation : ARRAY [1..4] OF BOOL;
	axEmergencyStopCabinet : ARRAY [1..2] OF BOOL;
	axDoorLocked : ARRAY [1..4] OF BOOL;
	axDoorUnlockDemand : ARRAY [1..4] OF BOOL;
	axDoorSeenUnlocked : ARRAY [1..4] OF BOOL;
	artDoorButton : ARRAY [1..4] OF R_TRIG;
	rtSafetyRelayReset : R_TRIG;
	tpSafetyRelayReset : TP;
	rtCellStart : R_TRIG;
	rtCellStop : R_TRIG;
	rtCellReset : R_TRIG;
	xEmergencyStopMpg : BOOL;
	xPhaseRelayOk : BOOL;
	xPressureRelayOk : BOOL;
	xSafetyRelayOk : BOOL;
	dwLiveFaultMask : DWORD;
	uiDoor : UINT;
	uiMagazine : UINT;
END_VAR
VAR CONSTANT
	ERR_ESTOP_STATION_1 : DWORD := DWORD#16#0000_0001;
	ERR_ESTOP_STATION_2 : DWORD := DWORD#16#0000_0002;
	ERR_ESTOP_STATION_3 : DWORD := DWORD#16#0000_0004;
	ERR_ESTOP_STATION_4 : DWORD := DWORD#16#0000_0008;
	ERR_ESTOP_CABINET_FRONT : DWORD := DWORD#16#0000_0010;
	ERR_ESTOP_CABINET_REAR  : DWORD := DWORD#16#0000_0020;
	ERR_ESTOP_MPG      : DWORD := DWORD#16#0000_0040;
	ERR_PHASE_RELAY    : DWORD := DWORD#16#0000_0080;
	ERR_PRESSURE_RELAY : DWORD := DWORD#16#0000_0100;
	ERR_SAFETY_RELAY   : DWORD := DWORD#16#0000_0200;
	ERR_DOOR_1_UNLOCKED : DWORD := DWORD#16#0000_0400;
	ERR_DOOR_2_UNLOCKED : DWORD := DWORD#16#0000_0800;
	ERR_DOOR_3_UNLOCKED : DWORD := DWORD#16#0000_1000;
	ERR_DOOR_4_UNLOCKED : DWORD := DWORD#16#0000_2000;
	WRN_SAFETY_RESET_REJECTED : UINT := UINT#1;
	WRN_DOOR_1_UNLOCK_REJECTED : UINT := UINT#2;
END_VAR

// --- BEGIN IMPLEMENTATION ---

fbFaultInjector(Request := FaultRequest);
FaultStatus := fbFaultInjector.Status;

FOR uiDoor := UINT#1 TO UINT#4 DO
	axEmergencyStopStation[uiDoor] := axEmergencyStopButtonStationInput[uiDoor]
		OR fbFaultInjector.axEmergencyStopStation[uiDoor];
	axDoorLocked[uiDoor] := axDoorLockClosedInput[uiDoor]
		AND NOT fbFaultInjector.axDoorUnlocked[uiDoor];
	artDoorButton[uiDoor](CLK := axDoorUnlockButtonInput[uiDoor]);

	IF uiDoor <= UINT#2 THEN
		uiMagazine := UINT#1;
	ELSE
		uiMagazine := UINT#2;
	END_IF;
	astEnclosureDoorStatus[uiDoor].xUnlockAllowed := NOT astMagazineStatus[uiMagazine].xEnabled AND NOT axMagazineMechanismBusy[uiMagazine];
	axDoorButtonLampOutput[uiDoor] := astEnclosureDoorStatus[uiDoor].xUnlockAllowed;

	IF artDoorButton[uiDoor].Q THEN
		IF astEnclosureDoorStatus[uiDoor].xUnlockAllowed THEN
			axDoorUnlockDemand[uiDoor] := TRUE;
			axDoorSeenUnlocked[uiDoor] := FALSE;
		ELSE
			RaiseWarning(uiCode := WRN_DOOR_1_UNLOCK_REJECTED + uiDoor - UINT#1);
		END_IF;
	END_IF;

	// Команда держится до фактического цикла «замок открылся -> снова закрылся».
	// Если магазин включили поверх открытого доступа, выход снимается немедленно.
	IF NOT astEnclosureDoorStatus[uiDoor].xUnlockAllowed THEN
		axDoorUnlockDemand[uiDoor] := FALSE;
		axDoorSeenUnlocked[uiDoor] := FALSE;
	ELSIF axDoorUnlockDemand[uiDoor] THEN
		IF NOT axDoorLocked[uiDoor] THEN
			axDoorSeenUnlocked[uiDoor] := TRUE;
		ELSIF axDoorSeenUnlocked[uiDoor] THEN
			axDoorUnlockDemand[uiDoor] := FALSE;
			axDoorSeenUnlocked[uiDoor] := FALSE;
		END_IF;
	END_IF;

	axDoorUnlockOutput[uiDoor] := axDoorUnlockDemand[uiDoor];
	astEnclosureDoorStatus[uiDoor].xLocked := axDoorLocked[uiDoor];
	astEnclosureDoorStatus[uiDoor].xUnlockOutput := axDoorUnlockOutput[uiDoor];
	astButtonStationIoStatus[uiDoor].xEmergencyStopPressed := axEmergencyStopStation[uiDoor];
	astButtonStationIoStatus[uiDoor].xButtonPressed := axDoorUnlockButtonInput[uiDoor];
	astButtonStationIoStatus[uiDoor].xButtonLightOn := axDoorButtonLampOutput[uiDoor];
	Status.axEmergencyStopReleased[uiDoor] := NOT axEmergencyStopStation[uiDoor];
	Status.axDoorReady[uiDoor] := astEnclosureDoorStatus[uiDoor].xUnlockAllowed OR axDoorLocked[uiDoor];
	Status.axButtonStationPressed[uiDoor] := astButtonStationIoStatus[uiDoor].xButtonPressed;
	Status.axButtonStationLightOn[uiDoor] := astButtonStationIoStatus[uiDoor].xButtonLightOn;
END_FOR;

FOR uiDoor := UINT#1 TO UINT#2 DO
	axEmergencyStopCabinet[uiDoor] := axEmergencyStopCabinetInput[uiDoor]
		OR fbFaultInjector.axEmergencyStopCabinet[uiDoor];
	Status.axEmergencyStopReleased[uiDoor + UINT#4] := NOT axEmergencyStopCabinet[uiDoor];
END_FOR;
xEmergencyStopMpg := xEmergencyStopMpgInput OR fbFaultInjector.xEmergencyStopMpg;
Status.axEmergencyStopReleased[7] := NOT xEmergencyStopMpg;

xPhaseRelayOk := xPhaseRelayOkInput AND NOT fbFaultInjector.xPhaseRelayFault;
xPressureRelayOk := xPressureRelayOkInput AND NOT fbFaultInjector.xPressureRelayFault;
xSafetyRelayOk := xSafetyRelayOkInput AND NOT fbFaultInjector.xSafetyRelayFault;

rtSafetyRelayReset(CLK := xSafetyRelayReset);
Status.xSafetyRelayResetAllowed := NOT xSafetyRelayOk AND NOT tpSafetyRelayReset.Q;
IF rtSafetyRelayReset.Q AND NOT Status.xSafetyRelayResetAllowed THEN
	RaiseWarning(uiCode := WRN_SAFETY_RESET_REJECTED);
END_IF;
tpSafetyRelayReset(
	IN := rtSafetyRelayReset.Q AND Status.xSafetyRelayResetAllowed,
	PT := T#1S
);
// Разрешение проверяется на фронте команды; после запуска выдаём полный импульс 1 с.
xSafetyRelayResetOutput := tpSafetyRelayReset.Q;
Status.xSafetyRelayResetActive := xSafetyRelayResetOutput;

rtCellStart(CLK := xCellStartButtonInput);
rtCellStop(CLK := xCellStopButtonInput);
rtCellReset(CLK := xCellResetButtonInput);
xCellEnablePulse := rtCellStart.Q;
xCellDisablePulse := rtCellStop.Q;
xCellResetPulse := rtCellReset.Q;

stFrontControlCabinetIoStatus.xEmergencyStopPressed := axEmergencyStopCabinet[1];
stFrontControlCabinetIoStatus.xStartPressed := xCellStartButtonInput;
stFrontControlCabinetIoStatus.xStopPressed := xCellStopButtonInput;
stFrontControlCabinetIoStatus.xResetPressed := xCellResetButtonInput;
stRearControlCabinetIoStatus.xEmergencyStopPressed := axEmergencyStopCabinet[2];
stRearControlCabinetIoStatus.xStartPressed := FALSE;
stRearControlCabinetIoStatus.xStopPressed := FALSE;
stRearControlCabinetIoStatus.xResetPressed := FALSE;
stMpgIoStatus.xEmergencyStopPressed := xEmergencyStopMpg;
stMpgIoStatus.xAxisX := xMpgAxisXInput;
stMpgIoStatus.xAxisY := xMpgAxisYInput;
stMpgIoStatus.xAxisZ := xMpgAxisZInput;
stMpgIoStatus.xMultiplier1 := xMpgMultiplier1Input;
stMpgIoStatus.xMultiplier10 := xMpgMultiplier10Input;
stMpgIoStatus.xMultiplier100 := xMpgMultiplier100Input;

dwLiveFaultMask := DWORD#0;
IF axEmergencyStopStation[1] THEN dwLiveFaultMask := dwLiveFaultMask OR ERR_ESTOP_STATION_1; END_IF;
IF axEmergencyStopStation[2] THEN dwLiveFaultMask := dwLiveFaultMask OR ERR_ESTOP_STATION_2; END_IF;
IF axEmergencyStopStation[3] THEN dwLiveFaultMask := dwLiveFaultMask OR ERR_ESTOP_STATION_3; END_IF;
IF axEmergencyStopStation[4] THEN dwLiveFaultMask := dwLiveFaultMask OR ERR_ESTOP_STATION_4; END_IF;
IF axEmergencyStopCabinet[1] THEN dwLiveFaultMask := dwLiveFaultMask OR ERR_ESTOP_CABINET_FRONT; END_IF;
IF axEmergencyStopCabinet[2] THEN dwLiveFaultMask := dwLiveFaultMask OR ERR_ESTOP_CABINET_REAR; END_IF;
IF xEmergencyStopMpg THEN dwLiveFaultMask := dwLiveFaultMask OR ERR_ESTOP_MPG; END_IF;
IF NOT xPhaseRelayOk THEN dwLiveFaultMask := dwLiveFaultMask OR ERR_PHASE_RELAY; END_IF;
IF NOT xPressureRelayOk THEN dwLiveFaultMask := dwLiveFaultMask OR ERR_PRESSURE_RELAY; END_IF;
IF NOT xSafetyRelayOk THEN dwLiveFaultMask := dwLiveFaultMask OR ERR_SAFETY_RELAY; END_IF;
IF (astMagazineStatus[1].xEnabled OR axMagazineMechanismBusy[1]) AND NOT axDoorLocked[1] THEN dwLiveFaultMask := dwLiveFaultMask OR ERR_DOOR_1_UNLOCKED; END_IF;
IF (astMagazineStatus[1].xEnabled OR axMagazineMechanismBusy[1]) AND NOT axDoorLocked[2] THEN dwLiveFaultMask := dwLiveFaultMask OR ERR_DOOR_2_UNLOCKED; END_IF;
IF (astMagazineStatus[2].xEnabled OR axMagazineMechanismBusy[2]) AND NOT axDoorLocked[3] THEN dwLiveFaultMask := dwLiveFaultMask OR ERR_DOOR_3_UNLOCKED; END_IF;
IF (astMagazineStatus[2].xEnabled OR axMagazineMechanismBusy[2]) AND NOT axDoorLocked[4] THEN dwLiveFaultMask := dwLiveFaultMask OR ERR_DOOR_4_UNLOCKED; END_IF;

Error.dwErrorActive := dwLiveFaultMask;
Error.dwAlarmActive := dwLiveFaultMask;
IF dwLiveFaultMask <> DWORD#0 THEN
	Error.dwErrorLast := dwLiveFaultMask;
END_IF;
Status.xPhaseRelayOk := xPhaseRelayOk;
Status.xPressureRelayOk := xPressureRelayOk;
Status.xSafetyRelayOk := xSafetyRelayOk;
Status.xGlobalError := dwLiveFaultMask <> DWORD#0;
Status.xReady := NOT Status.xGlobalError;

(* ---- FB_CONTROLLER_DIAGNOSTICS.st ---- *)
FUNCTION_BLOCK FB_CONTROLLER_DIAGNOSTICS
VAR_INPUT
    Request : ST_CONTROLLER_WEB_REQUEST;
    udiNowMs : UDINT;
    xReset : BOOL;
    xResetWarnings : BOOL;
END_VAR
VAR_OUTPUT
    Status : ST_CONTROLLER_WEB_STATUS;
    stWarning : ST_WARNING_EVENT;
END_VAR
VAR CONSTANT
    CPU_APPLICATION_STOPPED : DWORD := DWORD#16#0100_0000; // CPU 5A, исторический бит 19:24.
    CPU_RUN_ALARM_MASK : DWORD := DWORD#16#FEFF_FFFF; // Все причины, кроме состояния STOP приложения.
END_VAR
VAR
    uliAgeMs : ULINT;
    udiLastFrameAtMs : UDINT;
    xFrameAccepted : BOOL;
    xHaveFreshFrame : BOOL;
    xCpuValid : BOOL;
    xModulesValid : BOOL;
    dwCpuCurrent1 : DWORD;
    dwCpuCurrent2 : DWORD;
    dwCpuStoppedCurrent : DWORD;
    dwModuleCurrent : DWORD;
    xMemoryCurrent : BOOL;
    dwNext1 : DWORD;
    dwNext2 : DWORD;
    dwNextModule : DWORD;
    xNewAlarm : BOOL;
    xNewMemory : BOOL;
    xCausesGone : BOOL;
END_VAR

// --- BEGIN IMPLEMENTATION ---

xFrameAccepted := FALSE;
xNewAlarm := FALSE;
xNewMemory := FALSE;
// В STOP этот FB не исполняется: 5A в доставленном пакете относится к прошлой
// остановке/загрузке, а не к аварии уже работающего приложения. Убираем только
// этот бит, в том числе из прежней защёлки при online change; остальные причины
// сохраняют GLOBAL_STOP и прежний порядок сброса. История STOP остаётся в gateway.
Status.dwCpuAlarm1 := Status.dwCpuAlarm1 AND CPU_RUN_ALARM_MASK;
IF (Request.udiSequence <> UDINT#0) AND (Request.udiSequence <> Status.udiAckSeq) THEN
    // История обнаружений доставляется и после STOP; свежесть текущей нормы
    // проверяется отдельно и не следует из одного факта получения пакета.
    dwNext1 := (Status.dwCpuAlarm1 OR Request.dwCpuObserved1 OR Request.dwCpuCurrent1) AND CPU_RUN_ALARM_MASK;
    dwNext2 := Status.dwCpuAlarm2 OR Request.dwCpuObserved2 OR Request.dwCpuCurrent2;
    dwNextModule := Status.dwModuleAlarm OR Request.dwModuleObserved OR Request.dwModuleCurrent;
    xNewAlarm := (dwNext1 <> Status.dwCpuAlarm1) OR (dwNext2 <> Status.dwCpuAlarm2)
        OR (dwNextModule <> Status.dwModuleAlarm);
    Status.dwCpuAlarm1 := dwNext1;
    Status.dwCpuAlarm2 := dwNext2;
    Status.dwModuleAlarm := dwNextModule;
    xNewMemory := NOT Status.xMemoryWarning AND (Request.xMemoryObserved OR Request.xMemoryCurrent);
    IF xNewMemory THEN
        Status.xMemoryWarning := TRUE;
        stWarning.uiCode := UINT#1;
        stWarning.udiSequence := stWarning.udiSequence + UDINT#1;
        IF stWarning.udiSequence = UDINT#0 THEN stWarning.udiSequence := UDINT#1; END_IF;
    END_IF;

    IF udiNowMs >= Request.udiIssuedAtMs THEN
        uliAgeMs := UDINT_TO_ULINT(udiNowMs) - UDINT_TO_ULINT(Request.udiIssuedAtMs);
    ELSE
        uliAgeMs := ULINT#4294967296 + UDINT_TO_ULINT(udiNowMs) - UDINT_TO_ULINT(Request.udiIssuedAtMs);
    END_IF;
    xFrameAccepted := uliAgeMs <= ULINT#3000;
    xHaveFreshFrame := xFrameAccepted;
    IF xFrameAccepted THEN udiLastFrameAtMs := Request.udiIssuedAtMs; END_IF;
    // Кешированный 5A также не подтверждает восстановление настоящей аварии CPU.
    dwCpuStoppedCurrent := Request.dwCpuCurrent1 AND CPU_APPLICATION_STOPPED;
    xCpuValid := xFrameAccepted AND Request.xCpuValid AND (dwCpuStoppedCurrent = DWORD#0);
    xModulesValid := xFrameAccepted AND Request.xModulesValid;
    dwCpuCurrent1 := Request.dwCpuCurrent1;
    dwCpuCurrent2 := Request.dwCpuCurrent2;
    dwModuleCurrent := Request.dwModuleCurrent;
    xMemoryCurrent := Request.xMemoryCurrent;
    Status.udiAckSeq := Request.udiSequence;
END_IF;

// Абсолютный возраст проверяется и в первом скане после STOP/паузы задачи.
IF udiNowMs >= udiLastFrameAtMs THEN
    uliAgeMs := UDINT_TO_ULINT(udiNowMs) - UDINT_TO_ULINT(udiLastFrameAtMs);
ELSE
    uliAgeMs := ULINT#4294967296 + UDINT_TO_ULINT(udiNowMs) - UDINT_TO_ULINT(udiLastFrameAtMs);
END_IF;
Status.xCpuFresh := xHaveFreshFrame AND (uliAgeMs <= ULINT#12000) AND xCpuValid;
Status.xModulesFresh := xHaveFreshFrame AND (uliAgeMs <= ULINT#12000) AND xModulesValid;
Status.xAlarmActive := (Status.dwCpuAlarm1 <> DWORD#0) OR (Status.dwCpuAlarm2 <> DWORD#0)
    OR (Status.dwModuleAlarm <> DWORD#0);
xCausesGone := (((Status.dwCpuAlarm1 = DWORD#0) AND (Status.dwCpuAlarm2 = DWORD#0))
        OR (Status.xCpuFresh AND (dwCpuCurrent1 = DWORD#0) AND (dwCpuCurrent2 = DWORD#0)))
    AND ((Status.dwModuleAlarm = DWORD#0) OR (Status.xModulesFresh AND (dwModuleCurrent = DWORD#0)));
Status.xResetAllowed := Status.xAlarmActive AND xCausesGone AND NOT xNewAlarm;
IF xReset AND Status.xResetAllowed THEN
    Status.dwCpuAlarm1 := DWORD#0;
    Status.dwCpuAlarm2 := DWORD#0;
    Status.dwModuleAlarm := DWORD#0;
    Status.xAlarmActive := FALSE;
    Status.xResetAllowed := FALSE;
END_IF;
Status.xWarningResetAllowed := Status.xMemoryWarning AND Status.xCpuFresh
    AND NOT xMemoryCurrent AND NOT xNewMemory;
IF xResetWarnings AND Status.xWarningResetAllowed THEN
    Status.xMemoryWarning := FALSE;
    Status.xWarningResetAllowed := FALSE;
END_IF;

// После подтверждённого исчезновения причин снимается вход зависимого Stop,
// чтобы владельцы разрешили общий Reset. Защёлки и запрет Auto остаются до Reset.
Status.xGlobalStopRequired := Status.xAlarmActive AND (NOT xCausesGone OR xNewAlarm);

(* ---- FB_DI_FILTER.st ---- *)
FUNCTION_BLOCK FB_DI_FILTER
VAR_INPUT
	xEnable : BOOL;
	xInput : BOOL;
	tRise : TIME := T#20MS; // Стабильный 0 -> 1
	tFall : TIME := T#20MS; // Стабильный 1 -> 0
END_VAR
VAR_OUTPUT
	xFiltered : BOOL;
END_VAR
VAR
	tonRise : TON;
	tonFall : TON;
END_VAR

// --- BEGIN IMPLEMENTATION ---

// Каждая смена направления сбрасывает противоположный таймер. Короткие
// выбросы не накапливаются. При нулевом времени уровень меняется в этом скане.
IF NOT xEnable THEN
	xFiltered := FALSE;
END_IF;
tonRise(IN := xEnable AND xInput AND NOT xFiltered, PT := tRise);
tonFall(IN := xEnable AND NOT xInput AND xFiltered, PT := tFall);
IF xEnable THEN
	IF xInput AND ((tRise = T#0MS) OR tonRise.Q) THEN
		xFiltered := TRUE;
	ELSIF NOT xInput AND ((tFall = T#0MS) OR tonFall.Q) THEN
		xFiltered := FALSE;
	END_IF;
END_IF;

(* ---- FB_GEOMETRY_CONTROL.st ---- *)
FUNCTION_BLOCK FB_GEOMETRY_CONTROL
VAR_INPUT
	xInitialize : BOOL;
	uiAction : UINT;
	xSupported : BOOL;
	xSimulation : BOOL;
	xGlobalError : BOOL;
	xManual : BOOL;
	xCellRunning : BOOL;
	xRobotBusy : BOOL;
	xMotionBusy : BOOL;
	xHmiAlive : BOOL;
	xIoManual : BOOL;
	xReset : BOOL;
	xDriveAlarm : BOOL;
	xDriveRunning : BOOL;
	xPartAtEnd : BOOL;
	rSimulationTravel : REAL;
	Signals : ST_GEOMETRY_SIGNALS;
	Config : ST_GEOMETRY_CONFIG;
	tTransport : TIME;
	tFeedback : TIME;
	tResetPulse : TIME;
	uiTimeFactor : UINT := UINT#1;
END_VAR
VAR_IN_OUT
	Memory : ST_GEOMETRY_MEMORY;
END_VAR
VAR_OUTPUT
	Status : ST_GEOMETRY_STATUS;
	Warning : ST_WARNING_EVENT;
	xRunOutput : BOOL;
	xResetOutput : BOOL;
	xCommandAccepted : BOOL;
	xSimulationEmptyConfirmed : BOOL; // Одноцикловое принятое изъятие/подтверждение пустоты виртуальной ленты
END_VAR
VAR
	xInitialized : BOOL;
	xEnabled : BOOL;
	xReserved : BOOL;
	xTransport : BOOL;
	xManualRun : BOOL;
	xDisablePending : BOOL;
	xStopPending : BOOL;
	xEnableWanted : BOOL;
	xResetBusy : BOOL;
	xResetSeen : BOOL;
	xConfigurationValid : BOOL;
	xManualBase : BOOL;
	xCommandRejected : BOOL;
	dwControlBlockers : DWORD;
	tTransportScaled : TIME;
	tFeedbackScaled : TIME;
	tonTransport : TON;
	tonFeedback : TON;
	tonRemoved : TON;
	tonReset : TON;
	stRemoved : ST_GEOMETRY_CALL;
END_VAR

// --- BEGIN IMPLEMENTATION ---

IF xInitialize THEN xInitialized := FALSE; END_IF;
IF NOT xInitialized THEN
	// После рестарта конечный датчик не доказывает пустоту всей ленты.
	xEnabled := FALSE; xReserved := FALSE; xTransport := FALSE; xManualRun := FALSE;
	xDisablePending := FALSE; xStopPending := FALSE; xEnableWanted := FALSE; xResetBusy := FALSE; xResetSeen := FALSE;
	Memory.xRecoveryRequired := TRUE; xInitialized := TRUE;
END_IF;
xCommandAccepted := FALSE;
xSimulationEmptyConfirmed := FALSE;
xCommandRejected := FALSE;
xConfigurationValid := Config.xConfigured AND (Config.lrSpeedFactor >= 0.1)
	AND (Config.lrSpeedFactor <= 1.0) AND (Config.lrSafeZ < 0.0) AND (Config.lrSafeZ >= -10000.0);
tTransportScaled := UDINT_TO_TIME(MAX(UDINT#1, TIME_TO_UDINT(tTransport) / UINT_TO_UDINT(MAX(UINT#1, uiTimeFactor))));
tFeedbackScaled := UDINT_TO_TIME(MAX(UDINT#1, TIME_TO_UDINT(tFeedback) / UINT_TO_UDINT(MAX(UINT#1, uiTimeFactor))));

IF xDriveAlarm THEN Memory.dwAlarm := Memory.dwAlarm OR DWORD#1; END_IF;
IF Memory.dwAlarm <> DWORD#0 THEN
	Memory.xRecoveryRequired := TRUE;
	IF Signals.xRobotInteraction THEN Memory.xRobotStopLatched := TRUE; END_IF;
	xEnabled := FALSE; xEnableWanted := FALSE; xTransport := FALSE; xManualRun := FALSE;
	xDisablePending := FALSE; xStopPending := FALSE;
END_IF;
IF xGlobalError OR NOT xSupported OR xIoManual THEN
	IF Memory.xOccupied OR xReserved OR xTransport OR xManualRun THEN Memory.xRecoveryRequired := TRUE; END_IF;
	xEnabled := FALSE; xEnableWanted := FALSE; xTransport := FALSE; xManualRun := FALSE;
	xDisablePending := FALSE; xStopPending := FALSE;
	xResetBusy := FALSE;
END_IF;
IF NOT xHmiAlive OR NOT xManual OR xCellRunning THEN xManualRun := FALSE; END_IF;

IF Signals.xReserve AND xEnabled AND NOT xDisablePending AND NOT xStopPending
	AND xConfigurationValid AND NOT Memory.xOccupied
	AND NOT Memory.xRecoveryRequired AND NOT xPartAtEnd AND NOT xDriveRunning
	AND NOT xManualRun AND NOT xResetBusy AND NOT xGlobalError AND xSupported AND NOT xIoManual
	AND (Memory.dwAlarm = DWORD#0) THEN
	xReserved := TRUE; Memory.Part := Signals.Call;
END_IF;
IF Signals.xDeposited AND xReserved AND (Signals.Call.udiId <> UDINT#0)
	AND (Memory.udiLastDepositId <> Signals.Call.udiId) THEN
	Memory.xOccupied := TRUE; Memory.xAtEndSeen := FALSE;
	Memory.udiLastDepositId := Signals.Call.udiId;
	Memory.udiProducedPartsTotal := Memory.udiProducedPartsTotal + UDINT#1;
	Memory.Part := Signals.Call; Memory.Part.uiState := UINT#4;
	IF (Memory.Part.uiMachine >= UINT#1) AND (Memory.Part.uiMachine <= UINT#3) THEN
		GVL_GEOMETRY_CONTROL.astCalls[Memory.Part.uiMachine] := Memory.Part;
	END_IF;
	F_GEOMETRY_EVENT(Call := Memory.Part);
END_IF;
IF Signals.xReleased THEN
	xReserved := FALSE;
	// Штатное выключение завершает доставку; Stop запрещает пуск после отхода.
	IF Memory.xOccupied AND xEnabled AND NOT xStopPending AND NOT Memory.xRecoveryRequired
		AND (Memory.dwAlarm = DWORD#0) AND NOT xGlobalError THEN xTransport := TRUE; END_IF;
END_IF;

xManualBase := xSupported AND xManual AND NOT xCellRunning AND NOT xRobotBusy
	AND NOT xMotionBusy AND NOT Signals.xRobotInteraction AND NOT xReserved
	AND NOT xDisablePending AND NOT xStopPending
	AND xHmiAlive AND NOT xGlobalError AND NOT xIoManual AND NOT xResetBusy;
Status.xConfigAllowed := xManualBase AND NOT xEnabled AND NOT xDriveRunning AND NOT Memory.xOccupied;
// Допуск записи данных публикует RunGeometryControl независимо от состояния ГК.
// xConfigAllowed остаётся строгим допуском проверки с движением к базе.
// Включение и подтверждение пустоты зависят от выбранного ГК.
// Движение робота вне этой станции и работа ячейки не запрещают эти команды.
// Биты причин в astGeometryStatus: контракт описан в DOKS/24-geometry-control.md.
dwControlBlockers := DWORD#0;
IF NOT xSupported THEN dwControlBlockers := dwControlBlockers OR DWORD#1; END_IF;
IF NOT xHmiAlive THEN dwControlBlockers := dwControlBlockers OR DWORD#2; END_IF;
IF xGlobalError THEN dwControlBlockers := dwControlBlockers OR DWORD#4; END_IF;
IF xIoManual THEN dwControlBlockers := dwControlBlockers OR DWORD#8; END_IF;
IF Memory.dwAlarm <> DWORD#0 THEN dwControlBlockers := dwControlBlockers OR DWORD#16; END_IF;
IF Signals.xRobotInteraction THEN dwControlBlockers := dwControlBlockers OR DWORD#64; END_IF;
IF xReserved THEN dwControlBlockers := dwControlBlockers OR DWORD#128; END_IF;
IF xDriveRunning THEN dwControlBlockers := dwControlBlockers OR DWORD#256; END_IF;
IF xManualRun THEN dwControlBlockers := dwControlBlockers OR DWORD#512; END_IF;
IF xResetBusy THEN dwControlBlockers := dwControlBlockers OR DWORD#1024; END_IF;
IF xDisablePending OR xStopPending THEN dwControlBlockers := dwControlBlockers OR DWORD#2048; END_IF;
IF xTransport THEN dwControlBlockers := dwControlBlockers OR DWORD#8192; END_IF;
Status.dwEnableBlockers := dwControlBlockers;
IF NOT xConfigurationValid THEN Status.dwEnableBlockers := Status.dwEnableBlockers OR DWORD#32; END_IF;
IF xEnabled THEN Status.dwEnableBlockers := Status.dwEnableBlockers OR DWORD#4096; END_IF;
Status.xEnableAllowed := Status.dwEnableBlockers = DWORD#0;
Status.xDisableAllowed := xSupported AND (xEnabled OR xEnableWanted OR xDisablePending);
Status.dwConfirmBlockers := dwControlBlockers;
IF xEnableWanted AND NOT xConfigurationValid THEN Status.dwConfirmBlockers := Status.dwConfirmBlockers OR DWORD#32; END_IF;
IF NOT xEnableWanted AND NOT Memory.xRecoveryRequired THEN Status.dwConfirmBlockers := Status.dwConfirmBlockers OR DWORD#16384; END_IF;
IF xPartAtEnd THEN Status.dwConfirmBlockers := Status.dwConfirmBlockers OR DWORD#32768; END_IF;
Status.xConfirmAllowed := Status.dwConfirmBlockers = DWORD#0;
Status.xManualStartAllowed := xManualBase AND NOT xDriveAlarm AND (Memory.dwAlarm = DWORD#0) AND NOT xManualRun;
Status.xResetAllowed := (Memory.dwAlarm <> DWORD#0) AND NOT xResetBusy AND xSupported
	AND NOT xGlobalError AND NOT xIoManual
	AND NOT xRobotBusy AND NOT xMotionBusy AND NOT xManualRun AND NOT xTransport;
Status.xSimulationRemoveAllowed := xSimulation AND xSupported AND xHmiAlive
	AND NOT xGlobalError AND NOT xIoManual AND NOT xResetBusy
	AND Memory.xOccupied AND NOT Signals.xRobotInteraction AND NOT xReserved AND NOT xDriveRunning;

CASE uiAction OF
	UINT#1:
		IF Status.xEnableAllowed THEN
			IF Memory.xRecoveryRequired OR Memory.xOccupied OR xPartAtEnd THEN
				xEnableWanted := TRUE; Warning.uiCode := UINT#1; Warning.udiSequence := Warning.udiSequence + UDINT#1;
			ELSE xEnabled := TRUE; END_IF;
			xCommandAccepted := TRUE;
		END_IF;
	UINT#2:
		IF Status.xDisableAllowed THEN
			xEnableWanted := FALSE; xManualRun := FALSE;
			IF Signals.xRobotInteraction OR xReserved OR xTransport
			OR (Memory.xOccupied AND NOT Memory.xRecoveryRequired) THEN xDisablePending := TRUE;
			ELSE
				xEnabled := FALSE; xTransport := FALSE; xDisablePending := FALSE;
				IF Memory.xOccupied OR xReserved THEN Memory.xRecoveryRequired := TRUE; END_IF;
			END_IF;
			xCommandAccepted := TRUE;
		END_IF;
	UINT#3:
		IF Status.xConfirmAllowed THEN
			IF Memory.xOccupied AND (Memory.Part.udiId <> UDINT#0) THEN
				stRemoved := Memory.Part; stRemoved.uiState := UINT#8; F_GEOMETRY_EVENT(Call := stRemoved);
				IF (stRemoved.uiMachine >= UINT#1) AND (stRemoved.uiMachine <= UINT#3) THEN
					IF GVL_GEOMETRY_CONTROL.astCalls[stRemoved.uiMachine].udiId = stRemoved.udiId THEN
						GVL_GEOMETRY_CONTROL.astCalls[stRemoved.uiMachine] := stRemoved;
					END_IF;
				END_IF;
			END_IF;
			Memory.xOccupied := FALSE; Memory.xAtEndSeen := FALSE; Memory.xRecoveryRequired := FALSE;
			Memory.Part.udiId := UDINT#0; Memory.Part.uiMachine := UINT#0; Memory.Part.uiProductType := UINT#0;
			// Самостоятельное подтверждение состояния не включает станцию.
			xEnabled := xEnableWanted;
			xReserved := FALSE; xEnableWanted := FALSE; xCommandAccepted := TRUE;
			xSimulationEmptyConfirmed := xSimulation;
		END_IF;
	UINT#4:
		IF xEnableWanted OR Memory.xRecoveryRequired THEN
			xEnableWanted := FALSE; xEnabled := FALSE; xCommandAccepted := TRUE;
			Warning.uiCode := UINT#2; Warning.udiSequence := Warning.udiSequence + UDINT#1;
		END_IF;
	UINT#5:
		IF Status.xManualStartAllowed THEN
			xManualRun := TRUE; xCommandAccepted := TRUE;
			IF Memory.xOccupied THEN Memory.xRecoveryRequired := TRUE; xEnabled := FALSE; END_IF;
		END_IF;
	UINT#6:
		xManualRun := FALSE; xTransport := FALSE; xDisablePending := FALSE; xCommandAccepted := TRUE;
		IF Signals.xRobotInteraction OR xReserved THEN xStopPending := TRUE;
		ELSIF Memory.xOccupied THEN Memory.xRecoveryRequired := TRUE; xEnabled := FALSE; END_IF;
	UINT#7:
		IF Status.xSimulationRemoveAllowed THEN
			xCommandAccepted := TRUE; xSimulationEmptyConfirmed := TRUE;
			xTransport := FALSE; xManualRun := FALSE;
		END_IF;
END_CASE;
IF (uiAction >= UINT#1) AND (uiAction <= UINT#7) AND NOT xCommandAccepted THEN xCommandRejected := TRUE; END_IF;
IF xStopPending AND NOT Signals.xRobotInteraction THEN
	xEnabled := FALSE; xTransport := FALSE; xDisablePending := FALSE; xStopPending := FALSE;
	IF Memory.xOccupied OR xReserved THEN Memory.xRecoveryRequired := TRUE; END_IF;
END_IF;

// Сброс привода — настоящий импульс. Внутренняя авария снимается после импульса,
// только при исчезновении входа. Занятость и требование восстановления сохраняются.
IF xReset AND NOT xResetSeen AND Status.xResetAllowed THEN xResetBusy := TRUE; END_IF;
xResetSeen := xReset;
tonReset(IN := xResetBusy, PT := tResetPulse);
xResetOutput := xResetBusy AND NOT tonReset.Q AND xSupported AND NOT xIoManual AND NOT xGlobalError;
IF xResetBusy AND tonReset.Q THEN
	xResetBusy := FALSE;
	IF NOT xDriveAlarm AND NOT xDriveRunning THEN Memory.dwAlarm := DWORD#0; Memory.xRobotStopLatched := FALSE; END_IF;
END_IF;

IF xTransport AND xPartAtEnd THEN
	Memory.xAtEndSeen := TRUE; xTransport := FALSE;
END_IF;
// В ручном режиме датчик никогда не останавливает привод.
xRunOutput := (xTransport OR xManualRun) AND NOT Signals.xRobotInteraction
	AND NOT xGlobalError AND xSupported AND NOT xIoManual AND NOT xDriveAlarm
	AND (Memory.dwAlarm = DWORD#0) AND NOT xResetBusy;
tonTransport(IN := xTransport AND xRunOutput, PT := tTransportScaled);
tonFeedback(IN := (xRunOutput <> xDriveRunning) AND NOT xResetBusy AND xSupported AND NOT xIoManual AND NOT xGlobalError, PT := tFeedbackScaled);
IF tonTransport.Q THEN Memory.dwAlarm := Memory.dwAlarm OR DWORD#2; END_IF;
IF tonFeedback.Q THEN Memory.dwAlarm := Memory.dwAlarm OR DWORD#4; END_IF;
IF Memory.dwAlarm <> DWORD#0 THEN
	xEnabled := FALSE; xEnableWanted := FALSE; xRunOutput := FALSE;
	xDisablePending := FALSE; xStopPending := FALSE;
	xTransport := FALSE; xManualRun := FALSE; Memory.xRecoveryRequired := TRUE;
	IF Signals.xRobotInteraction THEN Memory.xRobotStopLatched := TRUE; END_IF;
END_IF;
// Выключаем только после подтверждённого конца доставки и останова привода.
// Освобождённый резерв без укладки не требует движения пустой ленты.
IF xDisablePending AND NOT Signals.xRobotInteraction AND NOT xReserved
	AND NOT xTransport AND NOT xManualRun AND NOT xDriveRunning AND NOT xResetBusy
	AND (NOT Memory.xOccupied OR Memory.xAtEndSeen) THEN
	xEnabled := FALSE; xDisablePending := FALSE;
END_IF;
tonRemoved(IN := Memory.xOccupied AND Memory.xAtEndSeen AND NOT xPartAtEnd
	AND NOT Memory.xRecoveryRequired AND NOT xTransport AND NOT xManualRun
	AND NOT xDriveRunning AND NOT xReserved AND NOT Signals.xRobotInteraction
	AND (Memory.dwAlarm = DWORD#0) AND NOT xGlobalError, PT := T#3S);
// Явное изъятие в SIMULATION подтверждает пустоту всей ленты сразу.
// В NORMAL освобождение по датчику по-прежнему требует непрерывные 3 секунды.
IF tonRemoved.Q OR (xSimulationEmptyConfirmed AND Memory.xOccupied) THEN
	stRemoved := Memory.Part; stRemoved.uiState := UINT#8; F_GEOMETRY_EVENT(Call := stRemoved);
	IF (stRemoved.uiMachine >= UINT#1) AND (stRemoved.uiMachine <= UINT#3) THEN
		IF GVL_GEOMETRY_CONTROL.astCalls[stRemoved.uiMachine].udiId = stRemoved.udiId THEN
			GVL_GEOMETRY_CONTROL.astCalls[stRemoved.uiMachine] := stRemoved;
		END_IF;
	END_IF;
	Memory.xOccupied := FALSE; Memory.xAtEndSeen := FALSE;
	Memory.Part.udiId := UDINT#0; Memory.Part.uiMachine := UINT#0; Memory.Part.uiProductType := UINT#0;
END_IF;
IF xPartAtEnd AND NOT xSimulationEmptyConfirmed AND NOT Memory.xOccupied AND NOT xReserved THEN
	Memory.xRecoveryRequired := TRUE; xEnabled := FALSE;
END_IF;
IF xCommandRejected THEN Warning.uiCode := UINT#3; Warning.udiSequence := Warning.udiSequence + UDINT#1; END_IF;
Status.xEnabled := xEnabled;
Status.xDisablePending := xDisablePending;
Status.xReserved := xReserved;
// Виртуальный датчик снимается моделью на следующем скане после принятой команды.
Status.xPartAtEnd := xPartAtEnd AND NOT xSimulationEmptyConfirmed;
Status.xOccupied := Memory.xOccupied OR xReserved OR Memory.xRecoveryRequired OR Status.xPartAtEnd;
Status.xPartStored := Memory.xOccupied;
Status.xReady := xEnabled AND xConfigurationValid AND NOT Status.xOccupied AND NOT xDriveRunning
	AND NOT xDisablePending AND NOT xStopPending
	AND (Memory.dwAlarm = DWORD#0) AND NOT xGlobalError AND xSupported AND NOT xIoManual AND NOT xResetBusy;
Status.xDriveRunning := xDriveRunning;
Status.xDriveAlarm := xDriveAlarm;
Status.xError := Memory.dwAlarm <> DWORD#0;
Status.xRobotStopRequired := Memory.xRobotStopLatched AND Status.xError;
Status.xResetBusy := xResetBusy;
Status.xConfirmationActive := xEnableWanted;
Status.xRecoveryRequired := Memory.xRecoveryRequired;
Status.xConfigured := xConfigurationValid;
Status.udiProducedPartsTotal := Memory.udiProducedPartsTotal;
Status.udiPartId := Memory.Part.udiId;
Status.uiMachine := Memory.Part.uiMachine;
Status.uiProductType := Memory.Part.uiProductType;
IF xSimulationEmptyConfirmed THEN Status.rTravel := REAL#0.0;
ELSIF xSimulation THEN Status.rTravel := rSimulationTravel;
ELSIF Memory.xAtEndSeen THEN Status.rTravel := REAL#1.0;
ELSIF xTransport THEN Status.rTravel := MIN(REAL#0.95, TIME_TO_REAL(tonTransport.ET) / TIME_TO_REAL(tTransportScaled));
ELSIF NOT Memory.xOccupied THEN Status.rTravel := REAL#0.0; END_IF;
IF Status.xError THEN Status.uiState := UINT#6;
ELSIF Memory.xRecoveryRequired THEN Status.uiState := UINT#5;
ELSIF xManualRun THEN Status.uiState := UINT#7;
ELSIF NOT xEnabled THEN Status.uiState := UINT#0;
ELSIF xReserved THEN Status.uiState := UINT#2;
ELSIF xTransport THEN Status.uiState := UINT#3;
ELSIF Memory.xOccupied THEN Status.uiState := UINT#4;
ELSE Status.uiState := UINT#1; END_IF;

(* ---- FB_GEOMETRY_CONTROL_SIMULATION.st ---- *)
FUNCTION_BLOCK FB_GEOMETRY_CONTROL_SIMULATION
VAR_INPUT
	xInitialize : BOOL;
	xRun : BOOL;
	xReset : BOOL;
	xDeposited : BOOL;
	udiPartId : UDINT;
	xRemove : BOOL;
	xAlarm : BOOL;
	uiTimeFactor : UINT := UINT#1;
	tTravel : TIME := T#6S;
END_VAR
VAR_OUTPUT
	xDriveRunning : BOOL;
	xDriveAlarm : BOOL;
	xPartAtEnd : BOOL;
	rTravel : REAL;
END_VAR
VAR
	xPart : BOOL;
	udiSeenDeposit : UDINT;
	udiPreviousClock : UDINT;
	udiDeltaMs : UDINT;
	rElapsedMs : REAL;
END_VAR

// --- BEGIN IMPLEMENTATION ---

IF xInitialize THEN
	xPart := FALSE; xPartAtEnd := FALSE; rTravel := REAL#0.0; udiSeenDeposit := UDINT#0;
	rElapsedMs := REAL#0.0; udiPreviousClock := GVL_HMI.udiHmiCommandClockMs;
END_IF;

// Накопленный путь сохраняется при останове и аварии. TON с IN=FALSE его теряет.
udiDeltaMs := MIN(UDINT#1000, GVL_HMI.udiHmiCommandClockMs - udiPreviousClock);
udiPreviousClock := GVL_HMI.udiHmiCommandClockMs;
IF xDeposited AND (udiPartId <> UDINT#0) AND (udiPartId <> udiSeenDeposit) THEN
	xPart := TRUE; xPartAtEnd := FALSE; rTravel := REAL#0.0; rElapsedMs := REAL#0.0; udiSeenDeposit := udiPartId;
END_IF;
IF xRemove THEN xPart := FALSE; xPartAtEnd := FALSE; rTravel := REAL#0.0; rElapsedMs := REAL#0.0; END_IF;
xDriveAlarm := xAlarm; // Сброс выхода не снимает удерживаемую физическую причину.
xDriveRunning := xRun AND NOT xDriveAlarm;
IF xPart AND NOT xPartAtEnd AND xDriveRunning THEN
	rElapsedMs := rElapsedMs + UDINT_TO_REAL(udiDeltaMs) * UINT_TO_REAL(MAX(UINT#1, uiTimeFactor));
	rTravel := MIN(REAL#1.0, rElapsedMs / MAX(REAL#1.0, TIME_TO_REAL(tTravel)));
	IF rTravel >= REAL#1.0 THEN xPartAtEnd := TRUE; END_IF;
END_IF;

(* ---- FB_GRIPPER_SIMULATION.st ---- *)
FUNCTION_BLOCK FB_GRIPPER_SIMULATION
VAR_INPUT
	xUsePhysicalFeedback : BOOL; // NORMAL SoftMotion: подтверждать реальные датчики
	xPhysicalIoReady : BOOL;
	PhysicalFeedback : ST_GRIPPER_STATUS;
	tPhysicalActionTimeout : TIME := T#10S;
	xTestInitialize : BOOL;
	auiTestContent : ARRAY [1..2] OF UINT;
	uiTestOrientation : UINT;
	xSimulationAccelerationEnable : BOOL; // Разрешить ускорение таймеров только в симуляции
	uiSimulationTimeFactor : UINT := 1; // Коэффициент виртуального времени 1..100
	Command : ST_GRIPPER_COMMAND; // Команда управления захватом
	FaultRequest : ST_GRIPPER_FAULT_REQUEST; // Единый контракт диагностической инъекции

    tGripper1OpenTime  : TIME := T#500MS; // Время открытия первого захвата
    tGripper1CloseTime : TIME := T#500MS; // Время закрытия первого захвата
    tGripper2OpenTime  : TIME := T#500MS; // Время открытия второго захвата
    tGripper2CloseTime : TIME := T#500MS; // Время закрытия второго захвата
    tRotateTime        : TIME := T#700MS; // Время смены рабочего захвата
END_VAR
VAR_OUTPUT
	Status : ST_GRIPPER_STATUS; // Рабочие статусы захвата
	Diag   : ST_GRIPPER_DIAG; // Состояние автомата и активное действие
	Error  : ST_GRIPPER_ERRORS; // Активные и последние ошибки
	FaultStatus : ST_FAULT_INJECTION_STATUS; // Состояние источника для HMI
END_VAR
VAR
	uiEffectiveTimeFactor : UINT;
	udiActionTime : UDINT;
	fbFaultInjector : FB_GRIPPER_FAULT_INJECTOR; // Изоляция тестовых источников от автомата
	eState        : E_GRIPPER_STATE := E_GRIPPER_STATE.IDLE; // Текущее состояние автомата захвата
    eActiveAction : E_ROBOT_ACTION := E_ROBOT_ACTION.NONE; // Выполняемое действие захвата

    tonAction      : TON; // Таймер выполнения действия
    xActionFault   : BOOL; // Неисправность, относящаяся к текущему действию
	xActionValid   : BOOL; // Получено допустимое действие захвата
    xActionRequired: BOOL; // Для действия требуется физическое переключение
    tActionTime    : TIME; // Нормативное время текущего действия
	xActionConfirmed : BOOL;
	xPhysicalGlobalFault : BOOL;
	xPhysicalGripper1Fault : BOOL;
	xPhysicalGripper2Fault : BOOL;
	xPhysicalRotationFault : BOOL;
    xInitialized   : BOOL; // Начальные состояния установлены
	rtReset         : R_TRIG; // Фронт команды сброса захвата
END_VAR
VAR CONSTANT
	ERR_GRIPPER_1   : DWORD := DWORD#16#0000_0001; // Ошибка первого захвата
    ERR_GRIPPER_2   : DWORD := DWORD#16#0000_0002; // Ошибка второго захвата
    ERR_GRIP_ROTATE : DWORD := DWORD#16#0000_0004; // Ошибка механизма поворота
    ERR_GRIP_ACTION : DWORD := DWORD#16#0000_0008; // Недопустимое действие захвата
    ERR_GRIP_GLOBAL : DWORD := DWORD#16#0000_0010; // Общая ошибка захвата
	WRN_RESET_EXECUTE_ACTIVE : UINT := 1; // Команда захвата ещё активна
	WRN_RESET_GLOBAL_FAULT   : UINT := 2; // Общая неисправность ещё активна
	WRN_RESET_GRIPPER_1_FAULT: UINT := 3; // Неисправность первого захвата ещё активна
	WRN_RESET_GRIPPER_2_FAULT: UINT := 4; // Неисправность второго захвата ещё активна
	WRN_RESET_ROTATION_FAULT : UINT := 5; // Неисправность поворота ещё активна
END_VAR

// --- BEGIN IMPLEMENTATION ---

uiEffectiveTimeFactor := uiSimulationTimeFactor;
IF NOT xSimulationAccelerationEnable THEN
	uiEffectiveTimeFactor := UINT#1;
ELSIF uiEffectiveTimeFactor < UINT#1 THEN
	uiEffectiveTimeFactor := UINT#1;
ELSIF uiEffectiveTimeFactor > UINT#100 THEN
	uiEffectiveTimeFactor := UINT#100;
END_IF;

IF NOT xInitialized THEN
    Status.xGripper1Open := TRUE;
    Status.xGripper1Closed := FALSE;

    Status.xGripper2Open := TRUE;
    Status.xGripper2Closed := FALSE;

    Status.xRotatedToBlank := TRUE;
    Status.xRotatedToDetail := FALSE;

    xInitialized := TRUE;
END_IF;

IF xTestInitialize THEN
	Status.xGripper1Open := auiTestContent[1] = UINT#0;
	Status.xGripper1Closed := NOT Status.xGripper1Open;
	Status.xGripper2Open := auiTestContent[2] = UINT#0;
	Status.xGripper2Closed := NOT Status.xGripper2Open;
	Status.xRotatedToBlank := uiTestOrientation = UINT#0;
	Status.xRotatedToDetail := NOT Status.xRotatedToBlank;
	eState := E_GRIPPER_STATE.IDLE;
	Error.dwErrorActive := DWORD#0;
END_IF;

// Не создаём подтверждение позиции по прошедшему времени в NORMAL.
IF xUsePhysicalFeedback THEN
	Status.xGripper1Open := PhysicalFeedback.xGripper1Open;
	Status.xGripper1Closed := PhysicalFeedback.xGripper1Closed;
	Status.xGripper2Open := PhysicalFeedback.xGripper2Open;
	Status.xGripper2Closed := PhysicalFeedback.xGripper2Closed;
	Status.xRotatedToBlank := PhysicalFeedback.xRotatedToBlank;
	Status.xRotatedToDetail := PhysicalFeedback.xRotatedToDetail;
END_IF;
xPhysicalGlobalFault := xUsePhysicalFeedback AND NOT xPhysicalIoReady;
xPhysicalGripper1Fault := xUsePhysicalFeedback AND Status.xGripper1Open AND Status.xGripper1Closed;
xPhysicalGripper2Fault := xUsePhysicalFeedback AND Status.xGripper2Open AND Status.xGripper2Closed;
xPhysicalRotationFault := xUsePhysicalFeedback AND Status.xRotatedToBlank AND Status.xRotatedToDetail;

// Ошибочная обратная связь блокирует владельца и до начала действия.
// Используем существующие биты GRIPPER и принятый эффект ROBOT_STOP.
IF xPhysicalGlobalFault THEN
	Error.dwErrorActive := Error.dwErrorActive OR ERR_GRIP_GLOBAL;
	eState := E_GRIPPER_STATE.ERROR;
END_IF;
IF xPhysicalGripper1Fault THEN
	Error.dwErrorActive := Error.dwErrorActive OR ERR_GRIPPER_1;
	eState := E_GRIPPER_STATE.ERROR;
END_IF;
IF xPhysicalGripper2Fault THEN
	Error.dwErrorActive := Error.dwErrorActive OR ERR_GRIPPER_2;
	eState := E_GRIPPER_STATE.ERROR;
END_IF;
IF xPhysicalRotationFault THEN
	Error.dwErrorActive := Error.dwErrorActive OR ERR_GRIP_ROTATE;
	eState := E_GRIPPER_STATE.ERROR;
END_IF;

rtReset(CLK := Command.xReset);

fbFaultInjector(
	Request := FaultRequest,
	eActiveAction := eActiveAction
);
FaultStatus := fbFaultInjector.Status;

IF rtReset.Q
AND (eState = E_GRIPPER_STATE.ERROR) THEN
	IF Command.xExecute THEN
		Diag.stWarning.uiCode := WRN_RESET_EXECUTE_ACTIVE;
	ELSIF fbFaultInjector.xGlobalFault OR xPhysicalGlobalFault THEN
		Diag.stWarning.uiCode := WRN_RESET_GLOBAL_FAULT;
	ELSIF fbFaultInjector.xGripper1Fault OR xPhysicalGripper1Fault THEN
		Diag.stWarning.uiCode := WRN_RESET_GRIPPER_1_FAULT;
	ELSIF fbFaultInjector.xGripper2Fault OR xPhysicalGripper2Fault THEN
		Diag.stWarning.uiCode := WRN_RESET_GRIPPER_2_FAULT;
	ELSIF fbFaultInjector.xRotationFault OR xPhysicalRotationFault THEN
		Diag.stWarning.uiCode := WRN_RESET_ROTATION_FAULT;
	ELSE
		Diag.stWarning.uiCode := UINT#0;
	END_IF;

	IF Diag.stWarning.uiCode <> UINT#0 THEN
		Diag.stWarning.udiSequence := Diag.stWarning.udiSequence + UDINT#1;
		IF Diag.stWarning.udiSequence = UDINT#0 THEN
			Diag.stWarning.udiSequence := UDINT#1;
		END_IF;
	END_IF;
END_IF;

xActionFault := fbFaultInjector.xActionFault;
xActionConfirmed := FALSE;
CASE eActiveAction OF
	E_ROBOT_ACTION.UNCLAMP_1:
		xActionConfirmed := Status.xGripper1Open AND NOT Status.xGripper1Closed;
		xActionFault := xActionFault OR xPhysicalGripper1Fault;
	E_ROBOT_ACTION.CLAMP_1:
		xActionConfirmed := Status.xGripper1Closed AND NOT Status.xGripper1Open;
		xActionFault := xActionFault OR xPhysicalGripper1Fault;
	E_ROBOT_ACTION.UNCLAMP_2:
		xActionConfirmed := Status.xGripper2Open AND NOT Status.xGripper2Closed;
		xActionFault := xActionFault OR xPhysicalGripper2Fault;
	E_ROBOT_ACTION.CLAMP_2:
		xActionConfirmed := Status.xGripper2Closed AND NOT Status.xGripper2Open;
		xActionFault := xActionFault OR xPhysicalGripper2Fault;
	E_ROBOT_ACTION.ROTATE_TO_BLANK:
		xActionConfirmed := Status.xRotatedToBlank AND NOT Status.xRotatedToDetail;
		xActionFault := xActionFault OR xPhysicalRotationFault;
	E_ROBOT_ACTION.ROTATE_TO_DETAIL:
		xActionConfirmed := Status.xRotatedToDetail AND NOT Status.xRotatedToBlank;
		xActionFault := xActionFault OR xPhysicalRotationFault;
END_CASE;
tActionTime := T#0S;

CASE eActiveAction OF
	E_ROBOT_ACTION.UNCLAMP_1:
		tActionTime := tGripper1OpenTime;
	E_ROBOT_ACTION.CLAMP_1:
		tActionTime := tGripper1CloseTime;
	E_ROBOT_ACTION.UNCLAMP_2:
		tActionTime := tGripper2OpenTime;
	E_ROBOT_ACTION.CLAMP_2:
		tActionTime := tGripper2CloseTime;
	E_ROBOT_ACTION.ROTATE_TO_BLANK,
	E_ROBOT_ACTION.ROTATE_TO_DETAIL:
		tActionTime := tRotateTime;

END_CASE;

	udiActionTime := TIME_TO_UDINT(tActionTime) / TO_UDINT(uiEffectiveTimeFactor);
	IF udiActionTime < UDINT#1 THEN
		udiActionTime := UDINT#1;
	END_IF;
	tActionTime := UDINT_TO_TIME(udiActionTime);

IF xUsePhysicalFeedback THEN
	tActionTime := tPhysicalActionTimeout;
END_IF;

tonAction(
    IN := (eState = E_GRIPPER_STATE.EXECUTE)
          AND NOT xActionFault
          AND NOT fbFaultInjector.xGlobalFault AND NOT xPhysicalGlobalFault,
    PT := tActionTime
);

CASE eState OF

    E_GRIPPER_STATE.IDLE:

        Status.xBusy := FALSE;
        Status.xDone := FALSE;
        Status.xError := FALSE;

        IF Command.xExecute THEN
            eActiveAction := Command.eAction;
			xActionValid := TRUE;
			xActionRequired := TRUE;

            CASE Command.eAction OF

				E_ROBOT_ACTION.UNCLAMP_1:
					xActionRequired := NOT (Status.xGripper1Open AND NOT Status.xGripper1Closed);

				E_ROBOT_ACTION.CLAMP_1:
					xActionRequired := NOT (Status.xGripper1Closed AND NOT Status.xGripper1Open);

				E_ROBOT_ACTION.UNCLAMP_2:
					xActionRequired := NOT (Status.xGripper2Open AND NOT Status.xGripper2Closed);

				E_ROBOT_ACTION.CLAMP_2:
					xActionRequired := NOT (Status.xGripper2Closed AND NOT Status.xGripper2Open);

				E_ROBOT_ACTION.ROTATE_TO_BLANK:
					xActionRequired := NOT (Status.xRotatedToBlank AND NOT Status.xRotatedToDetail);

				E_ROBOT_ACTION.ROTATE_TO_DETAIL:
					xActionRequired := NOT (Status.xRotatedToDetail AND NOT Status.xRotatedToBlank);

            ELSE
				xActionValid := FALSE;
                Error.dwErrorActive := Error.dwErrorActive OR ERR_GRIP_ACTION;
                eState := E_GRIPPER_STATE.ERROR;
            END_CASE;

			IF xActionValid THEN
				IF xActionRequired THEN
					eState := E_GRIPPER_STATE.EXECUTE;
				ELSE
					eState := E_GRIPPER_STATE.DONE;
				END_IF;
			END_IF;
        END_IF;

    E_GRIPPER_STATE.EXECUTE:

        Status.xBusy := TRUE;
        Status.xDone := FALSE;

		// Снятие Execute отменяет только незавершённое виртуальное действие и
		// сохраняет последнюю подтверждённую позицию захвата.
		IF NOT Command.xExecute THEN
			Status.xBusy := FALSE;
			eActiveAction := E_ROBOT_ACTION.NONE;
			eState := E_GRIPPER_STATE.IDLE;

		ELSIF fbFaultInjector.xGlobalFault OR xPhysicalGlobalFault THEN
            Error.dwErrorActive := Error.dwErrorActive OR ERR_GRIP_GLOBAL;
            eState := E_GRIPPER_STATE.ERROR;

        ELSIF xActionFault THEN

            CASE eActiveAction OF

                E_ROBOT_ACTION.UNCLAMP_1,
                E_ROBOT_ACTION.CLAMP_1:
                    Error.dwErrorActive := Error.dwErrorActive OR ERR_GRIPPER_1;

                E_ROBOT_ACTION.UNCLAMP_2,
                E_ROBOT_ACTION.CLAMP_2:
                    Error.dwErrorActive := Error.dwErrorActive OR ERR_GRIPPER_2;

                E_ROBOT_ACTION.ROTATE_TO_BLANK,
                E_ROBOT_ACTION.ROTATE_TO_DETAIL:
                    Error.dwErrorActive := Error.dwErrorActive OR ERR_GRIP_ROTATE;

            END_CASE;

            eState := E_GRIPPER_STATE.ERROR;

        ELSIF xUsePhysicalFeedback THEN
			IF xActionConfirmed THEN
				eState := E_GRIPPER_STATE.DONE;
			ELSIF tonAction.Q THEN
				CASE eActiveAction OF
					E_ROBOT_ACTION.UNCLAMP_1, E_ROBOT_ACTION.CLAMP_1:
						Error.dwErrorActive := Error.dwErrorActive OR ERR_GRIPPER_1;
					E_ROBOT_ACTION.UNCLAMP_2, E_ROBOT_ACTION.CLAMP_2:
						Error.dwErrorActive := Error.dwErrorActive OR ERR_GRIPPER_2;
					E_ROBOT_ACTION.ROTATE_TO_BLANK, E_ROBOT_ACTION.ROTATE_TO_DETAIL:
						Error.dwErrorActive := Error.dwErrorActive OR ERR_GRIP_ROTATE;
				END_CASE;
				eState := E_GRIPPER_STATE.ERROR;
			END_IF;

        ELSIF tonAction.Q THEN

            CASE eActiveAction OF

                E_ROBOT_ACTION.UNCLAMP_1:
                    Status.xGripper1Open := TRUE;
                    Status.xGripper1Closed := FALSE;

                E_ROBOT_ACTION.CLAMP_1:
                    Status.xGripper1Open := FALSE;
                    Status.xGripper1Closed := TRUE;

                E_ROBOT_ACTION.UNCLAMP_2:
                    Status.xGripper2Open := TRUE;
                    Status.xGripper2Closed := FALSE;

                E_ROBOT_ACTION.CLAMP_2:
                    Status.xGripper2Open := FALSE;
                    Status.xGripper2Closed := TRUE;

                E_ROBOT_ACTION.ROTATE_TO_BLANK:
                    Status.xRotatedToBlank := TRUE;
                    Status.xRotatedToDetail := FALSE;

                E_ROBOT_ACTION.ROTATE_TO_DETAIL:
                    Status.xRotatedToBlank := FALSE;
                    Status.xRotatedToDetail := TRUE;

            END_CASE;

            eState := E_GRIPPER_STATE.DONE;
        END_IF;

    E_GRIPPER_STATE.DONE:

        Status.xBusy := FALSE;
        Status.xDone := TRUE;

        IF NOT Command.xExecute THEN
            Status.xDone := FALSE;
            eActiveAction := E_ROBOT_ACTION.NONE;
            eState := E_GRIPPER_STATE.IDLE;
        END_IF;

    E_GRIPPER_STATE.ERROR:

        Status.xBusy := FALSE;
        Status.xDone := FALSE;
        Status.xError := TRUE;

        IF Command.xReset
        AND NOT Command.xExecute
        AND NOT fbFaultInjector.xGlobalFault
        AND NOT fbFaultInjector.xGripper1Fault
		AND NOT fbFaultInjector.xGripper2Fault
		AND NOT fbFaultInjector.xRotationFault
		AND NOT xPhysicalGlobalFault
		AND NOT xPhysicalGripper1Fault
		AND NOT xPhysicalGripper2Fault
		AND NOT xPhysicalRotationFault THEN

			Error.dwErrorLast := Error.dwErrorActive;
            Error.dwErrorActive := DWORD#0;
            Status.xError := FALSE;
            eActiveAction := E_ROBOT_ACTION.NONE;
            eState := E_GRIPPER_STATE.IDLE;
        END_IF;

END_CASE;

Diag.eState := eState;
Diag.eActiveAction := eActiveAction;

IF Error.dwErrorActive <> DWORD#0 THEN
	Error.dwErrorLast := Error.dwErrorActive;
END_IF;

Error.stErrorActive := UpdateErrorView(dwError := Error.dwErrorActive);
Error.stErrorLast := UpdateErrorView(dwError := Error.dwErrorLast);
Error.dwAlarmActive := Error.dwErrorActive;
FaultStatus.xResetAllowed := (Error.dwErrorActive <> DWORD#0)
	AND NOT FaultStatus.xActive
	AND NOT xPhysicalGlobalFault
	AND NOT xPhysicalGripper1Fault
	AND NOT xPhysicalGripper2Fault
	AND NOT xPhysicalRotationFault;
